(* IEC 61131-3 sources: daoli-st-library/DL_Algo (part 14) *)

(* ---- FB_DL_GainSchedPid.st ---- *)
(*
  组件名 Component   : FB_DL_GainSchedPid
  子库 Sublibrary    : DL_Algo
  版本 Version       : 1.0.0
  兼容性 Platform    : CODESYS 3.5 / TwinCAT 3 / 汇川 InoProShop / Machine Expert（仅 Standard.library）
  功能 Function      : 增益调度 PID（T0 标准语义件）：
                       1) 按调度变量 fSchedX 在断点表 afSchedX 上分区线性插值 Kc/Ti/Td 参数集；
                       2) 区间过渡加权平滑：插值参数经一阶惯性（tGainSmooth）再入 PID 核，
                          防分区切换瞬间增益阶跃引起执行器冲击；
                       3) 内嵌并行式 PID 核（P + I + D），积分钳位抗饱和，输出限幅；
                       4) 组态闸：断点数域 [2, 8]、断点严格递增、Ti > 0、增益非有限 → 故障锁存。
  边界 Boundary      : ① 本件只出控制量 fCtrlOut，不写物理 IO（由上层适配层承载）；
                       ② 除法防护：Ti 下限 1.0E-6 s、调度跨度判零、tCycle 域闸后再进算式；
                       ③ 非有限值（NaN 自反 + 无穷差值自减）判组态/输入非法，锁存安全侧；
                       ④ 调度变量越断点表两端时取端点参数（钳位外推禁止）；
                       ⑤ 故障锁存解除唯一路径 = bReset 上升沿（输入引脚，恒可达）；
                       ⑥ 无全局变量引用、无外部变量声明、无物理地址寻址。
  依赖 Depends       : Standard.library（R_TRIG）
  溯源 Origin        : IEC 61131-3 标准语义的道莅防御性实现（增益调度 + 并行 PID 均为
                       公开标准控制语义，T0 口径；参考 t2-5-modpid 参数域划分，零代码行复制）
  码位 Code          : 16#02_3_8C
  码表 Error codes（Algo 格 02_3_8C，单轨：故障 0x038C / 信息 0x028C）:
    16#0002_038C 故障级：组态非法（断点数越 [2,8] / 断点非严格递增 / Ti <= 0 /
                 参数非有限 / tCycle <= T#0S），锁存至 bReset 上升沿
    16#0002_028C 信息级：调度变量越端点已钳位（不置 bError，每拍瞬时口径）
  修订历史 Revision  :
    2026-11-19  v1.0.0  R44 首版（批次 1 · 序号 2）
*)

TYPE E_DL_GspState :
(
    eIdle  := 0,    // 空闲：未使能，出口冻结 / Idle, outputs frozen
    eRun   := 10,   // 运行：调度插值 + PID 闭环 / Running, scheduling plus PID loop
    eFault := 90    // 故障：组态非法锁存 / Fault, configuration latched
);
END_TYPE

FUNCTION_BLOCK FB_DL_GainSchedPid
VAR_INPUT
    bEnable    : BOOL;                        // 使能，FALSE 时出口冻结 [-] / Enable
    bReset     : BOOL;                        // 上升沿清故障锁存 [-] / Reset edge
    fSetpoint  : REAL;                        // 设定值 [工程单位] / Setpoint
    fFeedback  : REAL;                        // 反馈值 [工程单位] / Feedback
    fSchedX    : REAL;                        // 调度变量（工况量）[工程单位] / Scheduling variable
    afSchedX   : ARRAY[1..8] OF REAL;         // 断点表（须严格递增）[工程单位] / Scheduling breakpoints
    afKc       : ARRAY[1..8] OF REAL;         // 各断点比例增益 [无量纲] / Kc per breakpoint
    afTi       : ARRAY[1..8] OF REAL;         // 各断点积分时间 [秒] / Ti per breakpoint
    afTd       : ARRAY[1..8] OF REAL;         // 各断点微分时间 [秒] / Td per breakpoint
    nPtCount   : INT := 2;                    // 断点数 [个]，域 2..8 / Breakpoint count
    tGainSmooth: TIME := T#1S;                // 增益平滑惯性时间 [毫秒] / Gain smoothing lag
    fOutMin    : REAL := 0.0;                 // 输出下限 [%] / Output floor
    fOutMax    : REAL := 100.0;               // 输出上限 [%] / Output ceiling
    tCycle     : TIME := T#10MS;              // 扫描周期 [毫秒]，须与实际一致 / Scan cycle time
    bResetInt  : BOOL := TRUE;                // 使能下降沿后积分复归 [-] / Reset integral on disable
END_VAR
VAR_OUTPUT
    fCtrlOut   : REAL;                        // 控制量输出 [%] / Control output
    fKcUse     : REAL;                        // 平滑后生效比例增益 [无量纲] / Effective Kc
    fTiUse     : REAL;                        // 平滑后生效积分时间 [秒] / Effective Ti
    fTdUse     : REAL;                        // 平滑后生效微分时间 [秒] / Effective Td
    bError     : BOOL;                        // 故障锁存标志 [-] / Fault latch flag
    uErrId     : UDINT;                       // 事件码，0 = 无事件 / Event code
    eState     : E_DL_GspState;               // 状态出口，段尾单点映射 / State outlet
END_VAR
VAR
    rtReset    : R_TRIG;                      // 复位沿实例，段 0 每拍无条件刷新 / Reset edge
    _eState    : E_DL_GspState := E_DL_GspState.eIdle;  // 内部相位（CASE 唯一写入目标） / Internal phase
    _fErr      : REAL;                        // 偏差 [工程单位] / Error
    _fP        : REAL;                        // 比例项 [%] / Proportional term
    _fI        : REAL;                        // 积分项 [%] / Integral term
    _fD        : REAL;                        // 微分项 [%] / Derivative term
    _fErrPrev  : REAL;                        // 上拍偏差快照 [工程单位] / Previous error
    _fKcRaw    : REAL;                        // 插值比例增益 [无量纲] / Interpolated Kc
    _fTiRaw    : REAL;                        // 插值积分时间 [秒] / Interpolated Ti
    _fTdRaw    : REAL;                        // 插值微分时间 [秒] / Interpolated Td
    _fSeg      : REAL;                        // 插值段权重 [无量纲] / Interpolation weight
    _fCyS      : REAL;                        // 扫描周期秒值 [秒] / Cycle time in seconds
    _fSmK      : REAL;                        // 平滑系数 [无量纲] / Smoothing coefficient
    _nIdx      : INT;                         // 断点搜索索引 [-] / Breakpoint search index
    _bCfgBad   : BOOL;                        // 组态非法当拍量 [-] / Config illegal flag
    _bSchedClp : BOOL;                        // 调度钳位当拍量 [-] / Schedule clamped flag
    _fTiSafe   : REAL;                        // 积分时间安全值 [秒] / Ti safety value
END_VAR
VAR CONSTANT
    DL_PT_MAX  : INT   := 8;                  // 断点数上限，与数组维度一致 [个] / Breakpoint ceiling
    DL_PT_MIN  : INT   := 2;                  // 断点数下限 [个] / Breakpoint floor
    DL_MS_PER_S: REAL  := 1000.0;             // 毫秒 → 秒换算系数 [毫秒/秒] / Milliseconds per second
    DL_TI_MIN  : REAL  := 1.0E-6;             // 积分时间下限 [秒] / Ti floor
    DL_ABS_MAX : REAL  := 1.0E30;             // 有限值判定上界 [工程单位] / Finite value bound
    DL_EPS     : REAL  := 1.0E-9;             // 跨度判零容差 [工程单位] / Zero span tolerance
    DL_ZERO    : REAL  := 0.0;                // 零常量 [工程单位] / Zero constant
    DL_ONE     : REAL  := 1.0;                // 单位常量 [无量纲] / Unity constant
    DL_NO_TIME : TIME  := T#0S;               // 零时长哨兵 [毫秒] / Zero time sentinel
END_VAR

(* —— 段 0｜沿实例每拍无条件刷新（禁置于 IF/CASE 内） —— *)
rtReset(CLK := bReset);

(* —— 段 1｜瞬时量预清零（锁存量 _eState/积分项不入清单，禁同拍抹除） —— *)
_bCfgBad   := FALSE;
_bSchedClp := FALSE;
uErrId     := 16#0000_0000;

(* —— 段 2｜复位沿：故障一次性清干净，相位回空闲 —— *)
IF rtReset.Q THEN
    _eState  := E_DL_GspState.eIdle;
    _fI      := DL_ZERO;
    _fErrPrev:= DL_ZERO;
END_IF

(* —— 段 3｜周期换算与组态闸（覆盖全部参与换算引脚） —— *)
_fCyS := TIME_TO_REAL(tCycle) / DL_MS_PER_S;    // 毫秒 → 秒（TIME_TO_REAL 标准转换）
IF (tCycle = DL_NO_TIME) OR (nPtCount < DL_PT_MIN) OR (nPtCount > DL_PT_MAX) THEN
    _bCfgBad := TRUE;
END_IF
IF NOT _bCfgBad THEN
    _nIdx := 1;
    WHILE (_nIdx < nPtCount) AND (NOT _bCfgBad) DO
        IF (afSchedX[_nIdx] <> afSchedX[_nIdx]) OR (afKc[_nIdx] <> afKc[_nIdx])
           OR (afTi[_nIdx] <> afTi[_nIdx]) OR (afTd[_nIdx] <> afTd[_nIdx])
           OR (afSchedX[_nIdx + 1] <= afSchedX[_nIdx]) OR (afTi[_nIdx] <= DL_EPS)
           OR (afTi[_nIdx] > DL_ABS_MAX) THEN
            _bCfgBad := TRUE;               // 断点非递增 / 参数非有限 / Ti 无效
        END_IF
        _nIdx := _nIdx + 1;
    END_WHILE;
END_IF

(* —— 段 4｜主状态机：三态全覆盖 + ELSE 兜底 —— *)
CASE _eState OF

E_DL_GspState.eIdle:
    IF bEnable AND (NOT _bCfgBad) THEN
        _fI       := DL_ZERO;               // 入运行相前积分清零
        _fErrPrev := DL_ZERO;
        _eState   := E_DL_GspState.eRun;
    ELSIF bEnable AND _bCfgBad THEN
        bError    := TRUE;                  // 故障级配对置位（R45）
        uErrId    := 16#0002_038C;          // 组态非法锁存
        _eState   := E_DL_GspState.eFault;
    END_IF

E_DL_GspState.eRun:
    IF NOT bEnable THEN
        IF bResetInt THEN
            _fI := DL_ZERO;                 // 使能撤销按组态复归积分
        END_IF
        _eState := E_DL_GspState.eIdle;
    ELSE
        (* 调度插值：越端点钳位取端点参数并留信息码 *)
        IF fSchedX <= afSchedX[1] THEN
            _nIdx      := 1;
            _fSeg      := DL_ZERO;
            _bSchedClp := TRUE;
        ELSIF fSchedX >= afSchedX[nPtCount] THEN
            _nIdx      := nPtCount - 1;
            _fSeg      := DL_ONE;
            _bSchedClp := TRUE;
        ELSE
            _nIdx := 1;
            WHILE (_nIdx < nPtCount) AND (fSchedX >= afSchedX[_nIdx + 1]) DO
                _nIdx := _nIdx + 1;         // 断点严格递增已由组态闸保证
            END_WHILE;
            _fSeg := (fSchedX - afSchedX[_nIdx]) / (afSchedX[_nIdx + 1] - afSchedX[_nIdx]);
        END_IF
        _fKcRaw := afKc[_nIdx] + _fSeg * (afKc[_nIdx + 1] - afKc[_nIdx]);
        _fTiRaw := afTi[_nIdx] + _fSeg * (afTi[_nIdx + 1] - afTi[_nIdx]);
        _fTdRaw := afTd[_nIdx] + _fSeg * (afTd[_nIdx + 1] - afTd[_nIdx]);

        (* 一阶惯性平滑：系数域闸后加权，tGainSmooth 为零时直通 *)
        IF tGainSmooth <= DL_NO_TIME THEN
            _fSmK := DL_ONE;
        ELSE
            _fSmK := _fCyS / (_fCyS + TIME_TO_REAL(tGainSmooth) / DL_MS_PER_S);
        END_IF
        fKcUse := fKcUse + _fSmK * (_fKcRaw - fKcUse);
        fTiUse := fTiUse + _fSmK * (_fTiRaw - fTiUse);
        fTdUse := fTdUse + _fSmK * (_fTdRaw - fTdUse);
        IF _bSchedClp THEN
            uErrId := 16#0002_028C;         // 信息级：调度钳位（瞬时口径）
        END_IF

        (* PID 核：并行式，积分钳位抗饱和 *)
        _fErr := fSetpoint - fFeedback;
        _fP   := fKcUse * _fErr;
        _fTiSafe := MAX(fTiUse, DL_TI_MIN); // 积分时间下限护栏（除零前置）
        _fI := _fI + (fKcUse / _fTiSafe) * _fErr * _fCyS;
        _fD := (fKcUse * fTdUse / _fCyS) * (_fErr - _fErrPrev);
        fCtrlOut := _fP + _fI + _fD;
        IF fCtrlOut > fOutMax THEN
            fCtrlOut := fOutMax;
            _fI := _fI - (fKcUse / _fTiSafe) * _fErr * _fCyS;   // 上饱和积分回退
        ELSIF fCtrlOut < fOutMin THEN
            fCtrlOut := fOutMin;
            _fI := _fI - (fKcUse / _fTiSafe) * _fErr * _fCyS;   // 下饱和积分回退
        END_IF
        _fErrPrev := _fErr;
    END_IF

E_DL_GspState.eFault:
    ;                                   // 故障相驻留：出口冻结，只认复位沿（段 2 承载迁出）

ELSE
    bError := TRUE;                     // 兜底：非法相位锁存
    uErrId := 16#0002_038C;
    _eState := E_DL_GspState.eFault;
END_CASE

(* —— 段 5｜状态出口单点映射 —— *)
eState := _eState;
END_FUNCTION_BLOCK

(* ---- FB_DL_GainScheduler.st ---- *)
(*
    FB_DL_GainScheduler —— 分段增益调度
    ------------------------------------------------------------------
    分类      : DL_Algo / Control
    前缀      : FB_DL_
    版本      : 1.0.0
    溯源      : T2-5 Mod_PID（只借「参数域约束」的组织方式；源矩阵判定其参数域已取尽，
                仅剩「分段 / 手自动」这类手册细节，本件即分段这一侧的收口件）；
                迟滞判据、状态化输出、码位与分级 100% 自有；
                clean-room 重写，未复制任何闭源厂商源码，参考实现仅限 MIT/Apache 许可
    平台      : 纯 IEC 61131-3，CODESYS V3.5+ / TwinCAT 3 / InoProShop 通用
    作者      : 道莅代码库 · PLC编程专家（R18）
    ------------------------------------------------------------------
    功能说明  : 按调度变量（温度 / 流量 / 负载率）落在哪个断点区间，输出该段的一组
                Kp / Ki / Kd，解决「升温段要大 P、保温段要强 I」的分段整定需求；
                核心防御是边界迟滞：升段要越过「断点 + 迟滞半宽」，降段要跌破
                「断点 - 迟滞半宽」，杜绝边界抖动导致增益每拍来回跳；
                复位沿优先于定位，断点表严格递增在校验层一次性拦截；
                职责边界：本件只输出增益，不实现积分，也不做无扰切换——无扰由
                FB_DL_BumplessTransfer 与 PID 侧承担，避免与级联 PID 抢职责。
    错误码    : 16#0002_2301 调度变量非有限或变化被迟滞带抑制（保持当前段）——信息级，不置故障
                16#0002_2302 预留禁用（信息级，不得挪用）
                16#0002_2310 断点表非严格递增（非法组态）——故障级，输出保持末次并置故障
                16#0002_2311 段数越界（不在 2~4）——故障级，输出全 0 且不索引数组
                16#0002_2312 预留禁用（故障级，不得挪用）
    码位总账  : 16#0002_2301 用 / 16#0002_2302 预留 ｜ 16#0002_2310 用 / 16#0002_2311 用 / 16#0002_2312 预留
    状态机    : 无 CASE，段号由 uSeg 一个整数承载，非法状态由段数闸拦截，不可能出现
    采样约定  : fbTrigReset 在本体首部无条件刷新；本件无时间量，切换判定与任务周期无关，
                bSwitched 为单周期脉冲（每拍先清后置）。
    修订记录  : 2026-11-16 v1.0.0 首次入库（R18）
*)
FUNCTION_BLOCK FB_DL_GainScheduler
VAR_INPUT
    bEnable       : BOOL;                      // 使能，FALSE 输出保持末次并冻结段号 / enable, FALSE holds the last gains and freezes the segment
    bReset        : BOOL;                      // 复位，上升沿强制回到段 0 并清切换沿 / reset, rising edge forces segment zero and clears the switch pulse
    fScheduleVar  : REAL := 0.0;               // 调度变量（如温度）[用户单位] / scheduling variable such as temperature [user unit]
    afBreakpoint  : ARRAY[0..3] OF REAL;       // 分段上界断点，有效项 0~uSegCount-2，必须严格递增 [用户单位] / segment upper breakpoints, valid items 0~uSegCount-2, strictly increasing [user unit]
    afKp          : ARRAY[0..3] OF REAL;       // 各段比例增益 [无量纲] / proportional gain per segment [dimensionless]
    afKi          : ARRAY[0..3] OF REAL;       // 各段积分增益 [1/s] / integral gain per segment [1/s]
    afKd          : ARRAY[0..3] OF REAL;       // 各段微分增益 [s] / derivative gain per segment [s]
    uSegCount     : UINT := 2;                 // 段数 [段]，范围 2~4 / segment count [seg], range 2~4
    fHysteresis   : REAL := 0.5;               // 段边界迟滞带半宽 [用户单位]，范围 0.0~100.0，0 = 无迟滞 / half width of the boundary hysteresis band [user unit], range 0.0~100.0, 0 = none
END_VAR
VAR_OUTPUT
    fKp         : REAL;                        // 当前段比例增益 [无量纲] / proportional gain of the active segment [dimensionless]
    fKi         : REAL;                        // 当前段积分增益 [1/s] / integral gain of the active segment [1/s]
    fKd         : REAL;                        // 当前段微分增益 [s] / derivative gain of the active segment [s]
    uActiveSeg  : UINT;                        // 当前段号 0~3 [段] / active segment index 0~3 [seg]
    bSwitched   : BOOL;                        // 段切换单周期脉冲 / single-cycle segment switch pulse
    uSwitchCnt  : UDINT;                       // 累计切换次数，抖动监视用，饱和计数 [次] / accumulated switch count for chatter monitoring, saturating [times]
    eErr        : UDINT;                       // 错误码，0=正常 / error id, 0=ok
    bError      : BOOL;                        // 故障标志，eErr 为故障级时 TRUE / error flag, TRUE on fault-level eErr
END_VAR
VAR
    fbTrigReset : R_TRIG;                      // 复位沿检测实例，本体首部无条件刷新 / reset edge instance, refreshed unconditionally
    bInit       : BOOL := FALSE;               // 首扫标志，初值 FALSE，判据 NOT bInit / first-scan flag, initial FALSE, tested with NOT
    uSeg        : UINT;                        // 内部当前段号 [段] / internal active segment index [seg]
    uIdx        : UINT;                        // 断点遍历游标 [段] / breakpoint traversal cursor [seg]
    fHystEff    : REAL;                        // 生效迟滞半宽，钳位后使用 [用户单位] / effective hysteresis half width after clamping [user unit]
    bNonFin     : BOOL;                        // 调度变量非有限判定标志 / scheduling variable non-finite flag
    uSegLast    : UINT;                        // 上一拍段号，用于切换沿判定 [段] / previous cycle segment index for the switch edge [seg]
END_VAR
VAR CONSTANT
    DL_GS_SEG_MAX     : UINT := 4;             // 段数上限 [段] / segment count upper bound [seg]
    DL_GS_SEG_MIN     : UINT := 2;             // 段数下限 [段] / segment count lower bound [seg]
    DL_GS_LAST_IDX    : UINT := 3;             // 增益数组末索引 [段] / last gain array index [seg]
    DL_GS_HYST_MAX    : REAL := 100.0;         // 迟滞半宽上限 [用户单位] / hysteresis half width upper bound [user unit]
    DL_FLOAT_EPS      : REAL := 1.0E-6;        // 浮点判等容差 [用户单位] / float equality tolerance [user unit]
    DL_GS_INF_GUARD   : REAL := 4.0E38;        // 非有限幅值判定阈值 [用户单位] / non-finite magnitude guard [user unit]
    DL_GS_CNT_MAX     : UDINT := 16#FFFF_FFFE; // 切换计数饱和值 [次] / switch counter saturation value [times]
    DL_GS_ZERO        : REAL := 0.0;           // 零值常量，避免裸字面量 [无量纲] / zero constant, avoids a bare literal [dimensionless]
END_VAR

// 段 1｜边沿实例无条件周期刷新（红线：严禁放入条件分支）/ segment 1, unconditional edge refresh
fbTrigReset(CLK := bReset);

// 段 2｜输出与错误状态预置：bSwitched 每拍先清后置 / segment 2, preset outputs and error status
bSwitched := FALSE;                            // 单拍脉冲先清 / clear the single-cycle pulse first
eErr := 0;                                     // 预置无错误 / preset no error
bError := FALSE;                               // 预置无故障 / preset no fault

// 段 3｜首扫初始化（初值 FALSE，判据 NOT bInit）/ segment 3, first-scan initialisation
IF NOT bInit THEN
    uSeg := 0;                                 // 首扫落段 0 / start in segment zero
    uSegLast := 0;                             // 切换沿比较基准清零 / clear the switch edge reference
    uSwitchCnt := 0;                           // 切换计数清零 / clear the switch counter
    bInit := TRUE;                             // 首扫只做一次 / first scan runs once only
END_IF

// 段 4｜使能闸：失能保持末次增益并冻结段号 / segment 4, enable gate holds the last gains
IF NOT bEnable THEN
    uActiveSeg := uSeg;                        // 段号镜像保持 / keep the mirrored segment index
    RETURN;                                    // 失能即出口 / disabled is the exit
END_IF

// 段 5｜段数闸：越界即输出全 0 且不索引数组 / segment 5, segment count gate
IF (uSegCount < DL_GS_SEG_MIN) OR (uSegCount > DL_GS_SEG_MAX) THEN
    eErr := 16#0002_2311;                      // 段数越界故障码 / segment count out of range fault id
    bError := TRUE;                            // 置故障标志 / raise the error flag
    fKp := DL_GS_ZERO;                         // 输出全 0 / zero all gains
    fKi := DL_GS_ZERO;                         // 输出全 0 / zero the integral gain
    fKd := DL_GS_ZERO;                         // 输出全 0 / zero the derivative gain
    uActiveSeg := 0;                           // 段号回 0 / segment index back to zero
    RETURN;                                    // 故障级提前返回 / early return on fault
END_IF

// 段 6｜断点严格递增校验（浮点用大于号，禁用判等）/ segment 6, strict monotonic breakpoint check
FOR uIdx := 1 TO uSegCount - 2 DO
    IF NOT (afBreakpoint[uIdx] > afBreakpoint[uIdx - 1]) THEN
        eErr := 16#0002_2310;                  // 断点非法故障码 / illegal breakpoint fault id
        bError := TRUE;                        // 置故障标志 / raise the error flag
        uActiveSeg := uSeg;                    // 段号保持，输出保持末次 / keep the segment and the last gains
        RETURN;                                // 故障级提前返回 / early return on fault
    END_IF
END_FOR

// 段 7｜迟滞半宽双向钳位（负值视为无迟滞，超上限钳位）/ segment 7, hysteresis half width clamp
fHystEff := MIN(MAX(fHysteresis, DL_GS_ZERO), DL_GS_HYST_MAX); // 双侧钳位 / clamp both sides

// 段 8｜段号上界保护：段表缩短后旧段号可能越界 / segment 8, segment index upper bound protection
IF uSeg > (uSegCount - 1) THEN
    uSeg := uSegCount - 1;                     // 钳到最高段 / clamp to the highest segment
END_IF

// 段 9｜复位沿优先于定位 / segment 9, reset edge has priority over locating
IF fbTrigReset.Q THEN
    uSeg := 0;                                 // 强制回段 0 / force back to segment zero
END_IF

// 段 10｜迟滞定位：一次调用最多跨一段，跨多段交给后续拍 / segment 10, hysteresis locating, one step per cycle
bNonFin := (fScheduleVar <> fScheduleVar)
        OR (fScheduleVar > DL_GS_INF_GUARD)
        OR (fScheduleVar < -DL_GS_INF_GUARD);   // 非有限判定 / non-finite check
IF bNonFin THEN
    eErr := 16#0002_2301;                      // 非有限保持当前段（信息级不置故障）/ non-finite keeps the current segment, info level never raises a fault
ELSIF (NOT fbTrigReset.Q) THEN
    IF (uSeg < (uSegCount - 1)) AND (fScheduleVar > (afBreakpoint[uSeg] + fHystEff)) THEN
        uSeg := uSeg + 1;                      // 升段：必须越过断点加迟滞 / step up only beyond the breakpoint plus hysteresis
    ELSIF (uSeg > 0) AND (fScheduleVar < (afBreakpoint[uSeg - 1] - fHystEff)) THEN
        uSeg := uSeg - 1;                      // 降段：必须跌破断点减迟滞 / step down only below the breakpoint minus hysteresis
    END_IF
END_IF

// 段 11｜切换沿与抖动计数：段号变化才产生单拍脉冲 / segment 11, switch edge and chatter counting
IF uSeg <> uSegLast THEN
    bSwitched := TRUE;                         // 段号变化即置单拍脉冲 / raise the single-cycle pulse on any change
    IF uSwitchCnt < DL_GS_CNT_MAX THEN
        uSwitchCnt := uSwitchCnt + 1;          // 饱和加一，绝不回绕 / saturating increment, never wraps
    END_IF
END_IF
uSegLast := uSeg;                              // 记录本拍段号供下一拍比较 / remember this cycle segment for the next comparison

// 段 12｜增益输出：段号已由段 8 与段 5 双重保证在合法区间 / segment 12, publish the gains
fKp := afKp[uSeg];                             // 段号不超过 3，索引安全 / the segment index never exceeds three, indexing is safe
fKi := afKi[uSeg];                             // 积分增益取本段表值 / integral gain from the active segment row
fKd := afKd[uSeg];                             // 微分增益取本段表值 / derivative gain from the active segment row
uActiveSeg := uSeg;                            // 对外镜像段号 / publish the segment index
END_FUNCTION_BLOCK

(* ---- FB_DL_GapForceSwitchover.st ---- *)
(*==============================================================================
 * 组件名称 (Component)  : FB_DL_GapForceSwitchover
 * 所属子库 (Sublibrary) : DL_Algo
 * 当前版本 (Version)    : 1.0.0
 * 兼容性   (Platform)   : CODESYS 3.5+ / TwinCAT 3 / 汇川 InoProShop / 施耐德 Machine Expert
 *                         仅依赖 Standard.library（TON / R_TRIG / ABS / MAX），零厂商私有库
 * 功能描述 (Function)   : 压装/贴合类工步位置/压力双模式无扰切换：
 *                           eApproach 接近段：位置控趋近 fGapTargetMm，fCmdTrim = 间隙误差
 *                             修调（钳 ±fTrimMaxMm）；
 *                           接触判据：fForceN >= fContactN + 迟滞带 → eContact 过渡态，
 *                             冻结当时修调/速度作为衔接保持值（切换点速度不得突跳），
 *                             保持一个 tHoldXf 衔接窗后必迁出（单过渡态禁驻留，R285）；
 *                           eForceCtl 力控段：力偏差 → fForceTrimPct（钳 ±100%），
 *                             fCmdTrim 置 0；
 *                           tContactTmo 内未判接触 → eFault（eCause=eNoContact）；
 *                           力传感器非有限/超量程 → eFault（eCause=eForceBad）。
 * 接口     (Interface)  : 输入 fPosMm/fVelMmS 轴位姿、fForceN 力（N）、fContactN 接触判据
 *                         （N）、fGapTargetMm 目标间隙（mm）、fForceTargetN 力控目标（N）、
 *                         tContactTmo 接触超时、tHoldXf 衔接窗、fHysN 接触迟滞（N）、
 *                         fTrimMaxMm 修调限幅（mm）、fKpAppPct 接近修调增益（1/mm）、
 *                         fKpForcePct 力控增益（%/N）、fForceMaxN 力量程上限（N）、bReset；
 *                         输出 eMode 五态、fCmdTrim 位置环修调、fForceTrimPct 力环输出
 *                         （%）、eCause 成因、bError。
 * 边界     (Boundary)   : ① **属主边界（写死）：本件只出双模式状态与两侧修调量，不注入
 *                         轴指令、不接管压力环 PID**；修调限速可由上层用
 *                         `FB_DL_RateLimiter` 串联（本件不内嵌，规格依赖声明）。
 *                         ② 五态 CASE + ELSE 兜底 eFault（R6）；切换判据浮点容差比较
 *                         （迟滞带显式写出，禁 = 判等）。
 *                         ③ eContact 为单过渡态：tHoldXf 到时必迁 eForceCtl，禁驻留。
 *                         ④ 衔接保持值（_fTrimHold / _fVelHold）显式写出并在复位沿清零
 *                         （R311 预防：复位沿清状态与保持值）。
 *                         ⑤ 力超量程判据 = fForceN > fForceMaxN 或 fForceN < 0 或非有限
 *                         → eFault eForceBad（成因分码，R190 归因唯一）。
 *                         ⑥ 零全局耦合（无 GVL / VAR_EXTERNAL / 物理地址）。
 * 分工声明 (Scope)      : 与 `FB_DL_CoatingGapMeasure`（测量）与 `FB_DL_RollCompressForce-
 *                         Balance`（力平衡趋势）分工：切换闭环（本件）≠ 测量 ≠ 趋势。
 * 来源标签 (Source Tag) : T2-2 ◐（LBP 压机工艺分类只借"位置段/压力段"分类事实，切换器
 *                         实现自研）
 * 码表     (Codes)      : 本件不占用任何全局数字码位。出口为 ENUM 五态 + LREAL 组 +
 *                         ENUM 成因 + BOOL；数字码位待主控收口阶段统一派号。
 * 红线自检 (Redline)    : R1 ✓ 零 GVL/VAR_EXTERNAL ｜ R2 ✓ 零 %I/%Q/%M ｜ R3 ✓ 纯 IEC 61131-3
 *                         R4 ✓ 迟滞容差 + 非有限/超量程闸 + 修调钳位 ｜ R5 ✓ 声明逐行同行双语注释
 *                         R6 ✓ 五态 CASE 含 ELSE ｜ R7 ✓ 两 TON/一 R_TRIG 段 0 无条件刷新
 * 修订历史 (Revision)   : 2026-11-20  v1.0.0  R48 首版（批次 3 · 序号 13）
 *                         验收向量：接近段间隙误差修调；力越迟滞带 → eContact 冻结保持值；
 *                         衔接窗到 → eForceCtl；tContactTmo 无接触 → eFault eNoContact。
 *==============================================================================*)

TYPE E_DL_GfsMode :
(
    eIdle     := 0,    // 待机 / Idle
    eApproach := 10,   // 接近段（位置控）/ Approach phase, position control
    eContact  := 20,   // 接触过渡态（衔接保持，单过渡禁驻留）/ Contact transition, hold window
    eForceCtl := 30,   // 力控段 / Force control phase
    eFault    := 90    // 故障（等复位）/ Fault, awaiting reset
);
END_TYPE

TYPE E_DL_GfsCause :
(
    eNone       := 0,   // 无异常 / No anomaly
    eNoContact  := 1,   // 接近段超时未判接触 / No contact within timeout
    eForceBad   := 2,   // 力传感器非有限/超量程/负值 / Force sensor bad
    eCfgIllegal := 3,   // 组态非法 / Illegal configuration
    eModeBad    := 4    // 非法模式兜底 / Illegal mode fallback
);
END_TYPE

FUNCTION_BLOCK FB_DL_GapForceSwitchover
VAR_INPUT
    fPosMm      : LREAL := 0.0;    // 轴实际位置 [mm] / Axis actual position [mm]
    fVelMmS     : LREAL := 0.0;    // 轴实际速度 [mm/s] / Axis actual velocity [mm/s]
    fForceN     : LREAL := 0.0;    // 力/压力传感器实测 [N] / Force sensor measurement [N]
    fContactN   : LREAL := 5.0;    // 接触判据力，域 > 0 [N] / Contact force threshold [N]
    fGapTargetMm: LREAL := 0.0;    // 接近段目标间隙 [mm] / Approach target gap [mm]
    fForceTargetN: LREAL := 100.0; // 力控段目标力 [N] / Force-control target [N]
    tContactTmo : TIME := T#10S;   // 接近段接触超时，域 > T#0S [ms] / Contact timeout [ms]
    tHoldXf     : TIME := T#200MS; // eContact 衔接保持窗，域 > T#0S [ms] / Transition hold window [ms]
    fHysN       : LREAL := 0.5;    // 接触判据迟滞带，域 >= 0 [N] / Contact hysteresis band [N]
    fTrimMaxMm  : LREAL := 1.0;    // 位置环修调限幅，域 > 0 [mm] / Position trim limit [mm]
    fKpAppPct   : LREAL := 1.0;    // 接近段修调增益（间隙误差→修调） [1/mm] / Approach trim gain [1/mm]
    fKpForcePct : LREAL := 0.5;    // 力控段增益（力偏差→%） [%/N] / Force-control gain [%/N]
    fForceMaxN  : LREAL := 5000.0; // 力传感器量程上限，域 > fContactN [N] / Force range ceiling [N]
    bReset      : BOOL := FALSE;   // 故障复位，上升沿回 eIdle 并清保持值（R311） [-] / Fault reset, rising edge clears state and holds
END_VAR
VAR_OUTPUT
    eMode        : E_DL_GfsMode;   // 双模式状态出口 [-] / Mode state outlet
    fCmdTrim     : LREAL;          // 位置环速度/位置修调输出（力控段恒 0） [mm] / Position-loop trim outlet [mm]
    fForceTrimPct: LREAL;          // 力环修调输出（接近段恒 0） [%] / Force-loop trim outlet [%]
    eCause       : E_DL_GfsCause;  // 成因出口（锁存回放，R189） / Cause outlet, latched
    bError       : BOOL;           // 故障标志 [-] / Error flag
END_VAR
VAR
    _eMode     : E_DL_GfsMode := E_DL_GfsMode.eIdle;   // 内部状态（CASE 唯一写入目标） / Internal mode
    _eCause    : E_DL_GfsCause := E_DL_GfsCause.eNone; // 成因锁存量 / Latched cause
    _bFault    : BOOL;           // 故障锁存位（解除沿 = bReset 上升沿） / Latched fault bit
    _fTrimHold : LREAL := 0.0;   // 衔接保持值：接触瞬间修调 [mm] / Held trim at contact
    _fVelHold  : LREAL := 0.0;   // 衔接保持值：接触瞬间速度 [mm/s] / Held velocity at contact
    _fForceTrim: LREAL := 0.0;   // 力环修调锁存镜像 [%] / Force trim latch mirror
    _fCmdTrim  : LREAL := 0.0;   // 位置修调锁存镜像 [mm] / Position trim latch mirror
    _bErrScan  : BOOL;           // 力信号病当拍量（触发 eFault 用） / Force bad this scan
    _bNonFin   : BOOL;           // 输入非有限当拍量 [-] / Non-finite input this scan
    _bCfgBad   : BOOL;           // 组态非法当拍量 [-] / Illegal configuration this scan
    tonContactTmo: TON;          // 接近段接触超时定时器，段 0 无条件调用 / Contact timeout timer
    tonHoldXf  : TON;            // 衔接保持窗定时器，段 0 无条件调用 / Transition hold timer
    rtReset    : R_TRIG;         // 复位沿实例，段 0 无条件调用 / Reset edge instance
END_VAR
VAR CONSTANT
    DL_GFS_EPS   : LREAL := 1.0E-6;  // 浮点判零容差 [无量纲] / Float epsilon
    DL_GFS_ZERO  : LREAL := 0.0;     // 非有限差值判零基准 [-] / Non-finite difference zero base
    DL_GFS_PCTMAX: LREAL := 100.0;   // 力环修调行程上限 [%] / Force trim travel ceiling [%]
END_VAR

(* —— 段 0：非有限判 + 组态闸 + 两 TON 一沿无条件周期刷新 —— *)
_bNonFin := (fForceN <> fForceN) OR ((fForceN - fForceN) <> DL_GFS_ZERO)
         OR (fPosMm <> fPosMm) OR (fVelMmS <> fVelMmS);   // 力/位置/速度非有限（R245） / Non-finite force, position, velocity
_bCfgBad := (fContactN <= DL_GFS_ZERO) OR (fForceMaxN <= fContactN)
         OR (tContactTmo <= T#0S) OR (tHoldXf <= T#0S)
         OR (fTrimMaxMm <= DL_GFS_ZERO) OR (fHysN < DL_GFS_ZERO);   // 组态域闸 / Configuration gate
_bErrScan := _bNonFin OR (fForceN > fForceMaxN) OR (fForceN < DL_GFS_ZERO);   // 力信号病（超量程/负值/非有限） / Force signal bad
tonContactTmo(IN := (_eMode = E_DL_GfsMode.eApproach), PT := tContactTmo);   // 接触超时（进接近段计时，出段自复位） / Contact timeout
tonHoldXf(IN := (_eMode = E_DL_GfsMode.eContact), PT := tHoldXf);   // 衔接保持窗（进过渡态计时） / Transition hold window
rtReset(CLK := bReset);                                     // 复位沿，每拍必调 / Reset edge, every scan

(* —— 段 1：组态闸入故障 —— *)
IF _bCfgBad AND (NOT _bFault) THEN
    _bFault := TRUE;                                        // 组态非法锁存 / Latch config fault
    _eCause := E_DL_GfsCause.eCfgIllegal;                   // 归因：组态非法 / Cause: illegal config
    _eMode := E_DL_GfsMode.eFault;                          // 入故障态 / Enter fault
END_IF

(* —— 段 2：迁出链（复位沿：清状态与保持值，R311 预防） —— *)
IF rtReset.Q THEN
    _bFault := FALSE;                                       // 清故障锁存 / Clear fault latch
    _eCause := E_DL_GfsCause.eNone;                         // 清成因 / Clear cause
    _fTrimHold := 0.0;                                      // 清衔接保持修调 / Clear held trim
    _fVelHold := 0.0;                                       // 清衔接保持速度 / Clear held velocity
    _fCmdTrim := 0.0;                                       // 清修调镜像 / Clear trim mirror
    _fForceTrim := 0.0;                                     // 清力环镜像 / Clear force mirror
    _eMode := E_DL_GfsMode.eIdle;                           // 回待机 / Back to idle
END_IF

(* —— 段 3：力信号病 → 故障（成因分码 eForceBad，优先于时序） —— *)
IF _bErrScan AND (NOT _bFault) THEN
    _bFault := TRUE;                                        // 力信号病锁存 / Latch force fault
    _eCause := E_DL_GfsCause.eForceBad;                     // 归因：力传感器病 / Cause: force bad
    _eMode := E_DL_GfsMode.eFault;                          // 入故障态 / Enter fault
END_IF

(* —— 段 4：五态状态机（故障态由迁出链处理） —— *)
IF NOT _bFault THEN
    CASE _eMode OF

    E_DL_GfsMode.eIdle:
        _eMode := E_DL_GfsMode.eApproach;                   // 待机下一拍即入接近段（启动权交上层使能本件调用） / Idle proceeds to approach
        _fCmdTrim := 0.0;                                   // 修调清零起步 / Trim starts at zero

    E_DL_GfsMode.eApproach:
        _fCmdTrim := (fGapTargetMm - fPosMm) * fKpAppPct;   // 接近段修调 = 间隙误差×增益 / Approach trim from gap error
        IF _fCmdTrim > fTrimMaxMm THEN
            _fCmdTrim := fTrimMaxMm;                        // 修调上钳 / Clamp trim high
        ELSIF _fCmdTrim < -fTrimMaxMm THEN
            _fCmdTrim := -fTrimMaxMm;                       // 修调下钳 / Clamp trim low
        END_IF
        IF fForceN >= (fContactN + fHysN) THEN
            _fTrimHold := _fCmdTrim;                        // 接触瞬间冻结修调保持值（无扰衔接，头注释③） / Freeze trim at contact
            _fVelHold := fVelMmS;                           // 冻结接触瞬间速度（防切换突跳） / Freeze velocity at contact
            _fForceTrim := 0.0;                             // 力环修调起步零 / Force trim starts zero
            _eMode := E_DL_GfsMode.eContact;                // 越迟滞带上界：入接触过渡态 / Contact: enter transition
        ELSIF tonContactTmo.Q THEN
            _bFault := TRUE;                                // 超时未接触：故障锁存 / Timeout: latch fault
            _eCause := E_DL_GfsCause.eNoContact;            // 归因：未接触 / Cause: no contact
            _eMode := E_DL_GfsMode.eFault;                  // 入故障态 / Enter fault
        END_IF

    E_DL_GfsMode.eContact:
        _fCmdTrim := _fTrimHold;                            // 衔接窗内保持冻结修调（输出不突跳） / Hold frozen trim in window
        IF tonHoldXf.Q THEN
            _eMode := E_DL_GfsMode.eForceCtl;               // 衔接窗到必迁力控段（单过渡态禁驻留，R285） / Window done forces force phase
        END_IF

    E_DL_GfsMode.eForceCtl:
        _fCmdTrim := 0.0;                                   // 力控段位置修调归零 / Position trim zero in force phase
        _fForceTrim := (fForceTargetN - fForceN) * fKpForcePct;   // 力偏差 → 力环修调 / Force error to trim
        IF _fForceTrim > DL_GFS_PCTMAX THEN
            _fForceTrim := DL_GFS_PCTMAX;                   // 力环上钳 100% / Clamp force trim high
        ELSIF _fForceTrim < -DL_GFS_PCTMAX THEN
            _fForceTrim := -DL_GFS_PCTMAX;                  // 力环下钳 -100% / Clamp force trim low
        END_IF

    E_DL_GfsMode.eFault:
        ;                                                   // 故障态驻留：由段 2 迁出链复位处理 / Held by exit chain in stage 2

    ELSE
        _bFault := TRUE;                                    // 非法模式兜底（R6） / Illegal mode fallback
        _eCause := E_DL_GfsCause.eModeBad;                  // 归因：非法模式 / Cause: illegal mode
        _eMode := E_DL_GfsMode.eFault;                      // 强拉故障态 / Force fault

    END_CASE
END_IF

(* —— 段 5：出口单点映射（名实双出口同源，R191） —— *)
eMode := _eMode;                                            // 模式出口 / Mode outlet
fCmdTrim := _fCmdTrim;                                      // 位置修调出口（故障/待机零） / Position trim outlet
fForceTrimPct := _fForceTrim;                               // 力环修调出口 / Force trim outlet
eCause := _eCause;                                          // 成因出口 / Cause outlet
bError := _bFault OR _bCfgBad OR _bErrScan;                 // 故障标志三源合一 / Error flag
IF bError AND (NOT _bFault) THEN
    _bFault := TRUE;                                        // 当拍病亦锁存（防抖动复归） / Latch scan faults too
END_IF

END_FUNCTION_BLOCK

(* ---- FB_DL_GasDensityComp.st ---- *)
//==============================================================================
// 功能块：FB_DL_GasDensityComp ｜ 中文名称：反应釜气体密度温压补偿
// 所属子库：DL_Algo ｜ 版本：v1.0.0 ｜ 兼容：CODESYS V3.5+ / TwinCAT 3 / 汇川 InoProShop
// 功能描述：理想气体定律温压补偿——由工作温度与绝对压力换算气体密度：
//           rho = p·M / (R·T_K)，M 为介质摩尔质量 [g/mol]，R = 8.314462618
//           [J/(mol·K)]，T_K = T + 273.15。参考态密度 rho_ref 用参考温压
//           同式预计算（诊断出口）。骨架复用 FC_DL_AirDensity 的「域校验
//           + 钳位照算 + 非有限兜底」结构（该件介质常量固定为干空气/
//           水蒸气，反应釜介质摩尔质量可变，故本件以 M 引脚自持实现，
//           不调用该件——Algo 泳道内同口径双实现按 FC_DL_AirDensity 头
//           注释的零依赖纪律执行）。适用域：理想气体偏差可容忍的低压
//           工艺气（N2/Ar/H2/合成气等），近冷凝域给信息级外推提示。
// 开源溯源 (Origin)：道莅原创实现（参考理想气体状态方程与 FC_DL_AirDensity 域校验骨架 分类与参数域）
// 单位表：压力[千帕]（绝对）/ 温度[摄氏度] / 摩尔质量[克每摩尔] /
//         密度[千克每立方米] / 气体常数[J每摩尔开]
// 错误码表：16#0002_3201 信息级（温度/压力域外已钳位照算：温度域
//           [-40, 200] 摄氏度、压力域 [10, 2000] 千帕，不置 bError）/
//           16#0002_3202 信息级（理想气体外推提示：工作点温压比超出
//           参考态 0.5~2 倍温比或 10 倍压比工程带，按理想气体照算，
//           不置 bError）/ 16#0002_3205 预留禁用（不得挪用）/
//           16#0002_3210 故障级（摩尔质量 <= 0 或 > 200，或任一输入
//           非有限，组态非法，置 bError）/ 16#0002_3211 故障级（结果
//           非有限溢出，置 bError——该场景不可由 3210 的组态类判据
//           观测，属数值输出独立域）
// 状态机：E_DL_GasCompState（三态：eIdle=0 / eRun=10 / eFault=99），
//           CASE 含 ELSE 兜底，ELSE 置 3211 并冻结输出零
// 边界行为：① 摩尔质量域外或非有限 → 故障 3210 锁存，bReset 复位；
//           ② 温压域外 → 双侧钳位照算 + 信息 3201（现场宁要标注近似
//           的密度值，不因传感器越量程断链，与骨架件同策略）；
//           ③ 外推带 → 信息 3202 照算；④ 绝对温度下限 233.15 开由温度
//           下限保证，无除零面（T_K 恒正，R 为常量非零）；⑤ 未使能
//           输出冻结为零并 bValid := FALSE；⑥ 安全侧 = 故障/未使能路径
//           输出零密度，禁止残密度进入流量换算下游。
// 修订历史：v1.0.0 2026-11-17 首版（R24 派单 · ROADMAP P2 §670）
//==============================================================================

(*------------------------------------------------------------------------------
 * 枚举: E_DL_GasCompState（归属本功能块，同文件发布，全库唯一定义）
 * 含义: 补偿使能相位，每个成员在 CASE 中有且仅有一个标签。
 *-----------------------------------------------------------------------------*)
TYPE E_DL_GasCompState :
(
    eIdle  := 0,   // 空闲：未使能，输出冻结零 / Idle, not enabled, outputs frozen at zero
    eRun   := 10,  // 运行：使能且组态合法，每拍补偿 / Run, enabled with legal config, compensating per scan
    eFault := 99   // 故障：组态非法/非法状态 / Fault, illegal config or illegal state
);
END_TYPE

FUNCTION_BLOCK FB_DL_GasDensityComp
VAR_INPUT
    fPressKpa    : LREAL := 101.325;        // 工作绝对压力 [千帕]，域 10..2000，域外钳位照算 / Working absolute pressure [kPa], domain 10..2000
    fTempC       : LREAL := 20.0;           // 工作温度 [摄氏度]，域 -40..200，域外钳位照算 / Working temperature [degC], domain -40..200
    fMolarMassG  : LREAL := 28.96;          // 介质摩尔质量 [克每摩尔]，有效域 (0, 200]，空气 28.96 / Medium molar mass [g/mol], valid range (0, 200]
    fPressRefKpa : LREAL := 101.325;        // 参考态绝对压力 [千帕]，须 > 0 / Reference absolute pressure [kPa], must be > 0
    fTempRefC    : LREAL := 20.0;           // 参考态温度 [摄氏度]，须 > -273.15 / Reference temperature [degC], must be above absolute zero
    bEnable      : BOOL;                    // 补偿使能 [—] / Compensation enable
    bReset       : BOOL;                    // 故障复位 [—]，上升沿清组态锁存 / Fault reset, rising edge clears the config latch
END_VAR
VAR_OUTPUT
    fRhoKgM3     : LREAL;                   // 补偿密度 [千克每立方米] / Compensated density [kg/m3]
    fRhoRefKgM3  : LREAL;                   // 参考态密度（诊断出口）[千克每立方米] / Reference density, diagnostics outlet [kg/m3]
    eState       : E_DL_GasCompState;       // 补偿相位 [—] / Compensation phase
    eErr         : UDINT;                   // 错误码，0 = 无错，码位 16#0002_3201 起信息级、16#0002_3210 起故障级（分带见错误码表） / Error code, 0 = no error, band info/fault per the code table
    bError       : BOOL;                    // 故障级标志，仅故障级错误置位 / Fault-class flag, set only on fault-level codes
    bValid       : BOOL;                    // 输出可用标志 / Outputs usable flag
END_VAR
VAR
    _eState      : E_DL_GasCompState := E_DL_GasCompState.eIdle; // 当前相位 / Current phase
    _bParamBad   : BOOL;                    // 摩尔质量/参考态组态非法锁存 / Illegal molar mass or reference config latch
    _bInfoClamp  : BOOL;                    // 温压钳位信息当拍标志 / Temperature or pressure clamp info flag of this scan
    _bInfoExtrap : BOOL;                    // 外推带信息当拍标志 / Extrapolation-band info flag of this scan
    _fTUse       : LREAL;                   // 生效工作温度（已钳位）[摄氏度] / Effective working temperature, clamped
    _fPUse       : LREAL;                   // 生效工作压力（已钳位）[千帕] / Effective working pressure, clamped
    _fTKelvin    : LREAL;                   // 工作绝对温度 [开] / Working absolute temperature [K]
    _fTRefKelvin : LREAL;                   // 参考绝对温度 [开] / Reference absolute temperature [K]
    _bInit       : BOOL := FALSE;           // 首扫标志，初值 FALSE 取非判定 / First-scan flag, tested negated
    _bIllegal    : BOOL;                    // 非法状态标志 / Illegal state flag
END_VAR
VAR CONSTANT
    DL_GDC_R_UNIV  : LREAL := 8.314462618;  // 通用气体常数 [焦耳每摩尔开] / Universal gas constant [J/(mol K)]
    DL_GDC_KELVIN  : LREAL := 273.15;       // 摄氏转开尔文偏移 [开] / Celsius to Kelvin offset [K]
    DL_GDC_T_MIN   : LREAL := -40.0;        // 工作温度域下限 [摄氏度] / Working temperature domain floor [degC]
    DL_GDC_T_MAX   : LREAL := 200.0;        // 工作温度域上限 [摄氏度] / Working temperature domain ceiling [degC]
    DL_GDC_P_MIN   : LREAL := 10.0;         // 工作压力域下限 [千帕] / Working pressure domain floor [kPa]
    DL_GDC_P_MAX   : LREAL := 2000.0;       // 工作压力域上限 [千帕] / Working pressure domain ceiling [kPa]
    DL_GDC_M_MAX   : LREAL := 200.0;        // 摩尔质量域上限 [克每摩尔] / Molar mass domain ceiling [g/mol]
    DL_GDC_MRATIO  : LREAL := 10.0;         // 外推带压比门限 [倍] / Extrapolation pressure-ratio threshold [ratio]
    DL_GDC_TRATIO  : LREAL := 2.0;          // 外推带温比门限（双侧 0.5~2）[倍] / Extrapolation temperature-ratio threshold [ratio]
    DL_GDC_EPS     : LREAL := 1.0E-6;       // 浮点判零容差 [混合] / Float zero tolerance
    DL_GDC_INF     : LREAL := 1.7976931348623157E308; // LREAL 幅值上限 / LREAL magnitude ceiling
    DL_GDC_ZERO    : LREAL := 0.0;          // 零值常量，避免裸字面量 [混合] / Zero constant, avoids a bare literal
END_VAR

(*------------------------------------------------------------------------------
 * 段 1｜每拍预置：输出安全侧清零，单拍标志预清零
 *      Outputs cleared fail-safe first, one-shot flags pre-cleared
 *-----------------------------------------------------------------------------*)
fRhoKgM3    := DL_GDC_ZERO;              // 补偿密度先清（安全侧） / Compensated density cleared first
fRhoRefKgM3 := DL_GDC_ZERO;              // 参考密度先清 / Reference density cleared first
eErr   := 16#0000_0000;                  // 错误码每拍重算 / Error code recomputed
bError := FALSE;                         // 故障标志每拍重算 / Fault flag recomputed
bValid := FALSE;                         // 可用标志每拍重算 / Usable flag recomputed
_bInfoClamp  := FALSE;                   // 钳位信息预清零 / Clamp info pre-cleared
_bInfoExtrap := FALSE;                   // 外推信息预清零 / Extrapolation info pre-cleared
_bIllegal    := FALSE;                   // 非法状态预清零 / Illegal flag pre-cleared

(*------------------------------------------------------------------------------
 * 段 2｜首扫初始化
 *      First-scan initialisation
 *-----------------------------------------------------------------------------*)
IF NOT _bInit THEN
    _eState    := E_DL_GasCompState.eIdle; // 相位空闲起步 / Phase starts idle
    _bParamBad := FALSE;                   // 组态锁存清零 / Config latch cleared
    _bInit     := TRUE;                    // 首扫只做一次 / The first scan runs once
END_IF

(*------------------------------------------------------------------------------
 * 段 3｜组态防御闸：非有限（R79）+ 摩尔质量/参考态物理域
 *      Configuration defense gates: non-finite plus physical domains
 *-----------------------------------------------------------------------------*)
IF (fPressKpa <> fPressKpa) OR (ABS(fPressKpa) > DL_GDC_INF)
   OR (fTempC <> fTempC) OR (ABS(fTempC) > DL_GDC_INF)
   OR (fMolarMassG <> fMolarMassG) OR (ABS(fMolarMassG) > DL_GDC_INF)
   OR (fPressRefKpa <> fPressRefKpa) OR (ABS(fPressRefKpa) > DL_GDC_INF)
   OR (fTempRefC <> fTempRefC) OR (ABS(fTempRefC) > DL_GDC_INF) THEN
    _bParamBad := TRUE;                    // 非有限归组态非法锁存 / Non-finite folded into the config fault latch
END_IF
IF (NOT _bParamBad)
   AND ((fMolarMassG <= DL_GDC_EPS) OR (fMolarMassG > DL_GDC_M_MAX)
        OR (fPressRefKpa <= DL_GDC_EPS) OR (fTempRefC <= (-DL_GDC_KELVIN + 1.0))) THEN
    _bParamBad := TRUE;                    // 摩尔质量/参考态组态非法锁存 / Molar mass or reference config latched
END_IF
IF bReset THEN
    _bParamBad := FALSE;                   // 复位清组态锁存 / Reset clears the config latch
END_IF

(*------------------------------------------------------------------------------
 * 段 4｜相位机（CASE 含 ELSE 兜底；未使能/异常一律落故障态全零）
 *      Phase machine with ELSE fallback, not-enabled or anomaly to fault
 *-----------------------------------------------------------------------------*)
IF (NOT bEnable) OR _bParamBad THEN
    _eState := E_DL_GasCompState.eFault;   // 未使能或组态非法转故障态（全零） / Not enabled or illegal config, fault with zeros
ELSE
CASE _eState OF

    E_DL_GasCompState.eIdle:               // 空闲：使能即进运行
        IF bEnable THEN
            _eState := E_DL_GasCompState.eRun; // 进运行 / To run
        END_IF

    E_DL_GasCompState.eRun:                // 运行：每拍补偿（段 5 执行）
        IF NOT bEnable THEN
            _eState := E_DL_GasCompState.eFault; // 使能撤销转故障态（全零） / Enable dropped, fault with zeros
        END_IF

    E_DL_GasCompState.eFault:              // 故障：使能且复位沿回运行
        IF bEnable AND (NOT _bParamBad) THEN
            _eState := E_DL_GasCompState.eRun; // 回运行 / Back to run
        END_IF

    ELSE                                   // 非法状态兜底（R21：CASE 必带 ELSE）
        _bIllegal := TRUE;                 // 标记非法状态 / Flag the illegal state
        _eState   := E_DL_GasCompState.eFault; // 回故障态（全零） / Back to fault, zeros
END_CASE
END_IF

(*------------------------------------------------------------------------------
 * 段 5｜补偿计算（仅运行态）：域钳位照算 + 外推带提示 + 理想气体定律
 *      Compensation in the run phase: clamp-and-continue plus ideal-gas law
 *-----------------------------------------------------------------------------*)
IF _eState = E_DL_GasCompState.eRun THEN
    _fTUse := fTempC;                      // 工作温度生效 / Working temperature applied
    IF (_fTUse < DL_GDC_T_MIN) OR (_fTUse > DL_GDC_T_MAX) THEN
        _fTUse := MIN(MAX(_fTUse, DL_GDC_T_MIN), DL_GDC_T_MAX); // 温度双侧钳位 / Two-sided temperature clamp
        _bInfoClamp := TRUE;               // 钳位信息置位 / Clamp info raised
    END_IF
    _fPUse := fPressKpa;                   // 工作压力生效 / Working pressure applied
    IF (_fPUse < DL_GDC_P_MIN) OR (_fPUse > DL_GDC_P_MAX) THEN
        _fPUse := MIN(MAX(_fPUse, DL_GDC_P_MIN), DL_GDC_P_MAX); // 压力双侧钳位 / Two-sided pressure clamp
        _bInfoClamp := TRUE;               // 钳位信息置位 / Clamp info raised
    END_IF
    _fTKelvin    := _fTUse + DL_GDC_KELVIN;     // 工作绝对温度 [开]，下限 233.15 恒正 / Working Kelvin, floor 233.15, always positive
    _fTRefKelvin := fTempRefC + DL_GDC_KELVIN;  // 参考绝对温度 [开] / Reference Kelvin
    fRhoKgM3 := (_fPUse * 1000.0) * (fMolarMassG / 1000.0) / (DL_GDC_R_UNIV * _fTKelvin); // 理想气体密度 [千克每立方米]，分母恒正 / Ideal-gas density, denominator always positive
    fRhoRefKgM3 := (fPressRefKpa * 1000.0) * (fMolarMassG / 1000.0) / (DL_GDC_R_UNIV * _fTRefKelvin); // 参考态密度 [千克每立方米] / Reference density
    IF (_fPUse > DL_GDC_MRATIO * fPressRefKpa)
       OR (_fTKelvin < (0.5 * _fTRefKelvin)) OR (_fTKelvin > (DL_GDC_TRATIO * _fTRefKelvin)) THEN
        _bInfoExtrap := TRUE;              // 理想气体外推带提示（照算） / Extrapolation-band notice, computed as-is
    END_IF
END_IF

(*------------------------------------------------------------------------------
 * 段 6｜码位出口与放行（故障级码 3 行内置 bError，R45/R101 配对）
 *      Code outlet and release, fault codes paired with bError
 *-----------------------------------------------------------------------------*)
IF _bIllegal THEN
    eErr   := 16#0002_3211;                // 故障级：状态机兜底（结果域） / Fault: state machine fallback
    bError := TRUE;                        // 置故障标志 / Raise the fault flag
ELSIF _bParamBad THEN
    eErr   := 16#0002_3210;                // 故障级：组态非法 / Fault: illegal configuration
    bError := TRUE;                        // 置故障标志 / Raise the fault flag
ELSIF _bInfoClamp THEN
    eErr := 16#0002_3201;                  // 信息级：温压域外已钳位照算 / Info: clamped, computed as-is
ELSIF _bInfoExtrap THEN
    eErr := 16#0002_3202;                  // 信息级：理想气体外推带照算 / Info: extrapolation band, computed as-is
END_IF

bValid := (NOT bError) AND (_eState = E_DL_GasCompState.eRun); // 仅运行态放行 / Usable only in the run phase
eState := _eState;                       // 相位出口 / Phase outlet
END_FUNCTION_BLOCK

(* ---- FB_DL_GatedUpdateFilter.st ---- *)
(*==============================================================================
 * 组件名称 (Component)  : FB_DL_GatedUpdateFilter
 * 所属子库 (Sublibrary) : DL_Algo
 * 当前版本 (Version)    : 1.0.0
 * 兼容性   (Platform)   : CODESYS 3.5+ / TwinCAT 3 / 汇川 InoProShop / 施耐德 Machine Expert
 *                         仅依赖 Standard.library（TON），零厂商私有库
 * 功能描述 (Function)   : 门控更新滤波：**仅在允许窗口内采样，窗口外保持上次值**。
 *                         与低通 / 限速不同，本件不做任何数值整形，只决定「这一拍要不要采纳」，
 *                         因此阶跃与斜率在窗口内原样通过（无失真、无滞后）。
 *                         典型用途：剔除运动段/换型段的动态值、只在静止窗口内采重量、
 *                         只在保压阶段记录压力稳态值。
 *                         窗口外持续时长用 TON 累计；超过 tMaxHold 置 bStale=TRUE（信息级），
 *                         提示上游「数据已陈旧」，但**输出仍保持**（保持语义不变）。
 *                         恢复路径：bGate 重新为 TRUE 即回到新鲜；故障态由 bEnable 跌落或 bReset 解除。
 * 接口     (Interface)  : 输入 bEnable 使能、bReset 复位到当前输入、fIn 采样输入 [EU]、
 *                         bGate 窗口使能（TRUE = 本拍采纳）、tMaxHold 允许的最大保持时长 [s]；
 *                         输出 fOut 输出值 [EU]、bStale 数据是否陈旧、tHeldElapsed 已保持时长 [s]、
 *                         bValid 输出有效、bError、uErrorId。
 * 边界     (Boundary)   : ① 属主边界：只做门控与保持，不做平滑、不做离群剔除（另件）。
 *                         ② 非有限输入防御：窗口内（bGate=TRUE）遇非有限值 → 故障态 16#0006_0002，
 *                         输出冻结；窗口外（bGate=FALSE）不读取 fIn，故非有限值不判故障
 *                         （这是本件的语义：窗口外输入无意义）。
 *                         ③ tMaxHold < 0 钳到 T#0S 并置信息码 16#0006_0001；T#0S 表示不判陈旧
 *                         （bStale 恒 FALSE，TON 的 Q 仍按 PT=0 立即为真，故显式屏蔽）。
 *                         ④ **TON 无条件每周期调用**（R7），位于 CASE 之外。
 *                         ⑤ 零全局耦合（无 GVL / VAR_EXTERNAL / 物理地址）。
 * 分工声明 (Scope)      : 与 `FB_DL_HoldLastGoodFilter` 分工：坏值（判据失效）保持归那件、
 *                         时间窗门控归本件；与 `FB_DL_PeakHoldFilter` 分工：峰值保持归那件。
 * 来源标签 (Source Tag) : 原创实现（无外部代码引入）
 * 码表     (Codes)      : 16#0006_0000 无故障 / 16#0006_0001 保持时长非法已钳位（信息级）/
 *                         16#0006_0002 窗口内输入非有限（故障级）/ 16#0006_0005 非法状态（故障级）。
 * 红线自检 (Redline)    : R1 ✓ 零 GVL/VAR_EXTERNAL ｜ R2 ✓ 零 %I/%Q/%M ｜ R3 ✓ 纯 IEC 61131-3
 *                         R4 ✓ 非有限拒绝（仅窗口内）+ 时长域闸 + 无除法 ｜ R5 ✓ 声明逐行同行双语注释
 *                         R6 ✓ 四态 ENUM + CASE + ELSE 兜底 ｜ R7 ✓ TON 实例 CASE 外无条件刷新
 * 修订历史 (Revision)   : 2026-11-23  v1.0.0  R77 首版（批次 B3 · 序号 12）
 * 验收向量 (Acceptance) : ① bGate=TRUE 时 fIn 由 10 变 20 → 当拍 fOut=20；
 *                         ② 随后 bGate=FALSE 且 fIn=99 → fOut 保持 20（不采纳）, bStale=FALSE（未超时）；
 *                         ③ bGate 持续 FALSE 超过 tMaxHold=T#1S → bStale=TRUE，fOut 仍保持 20；
 *                         ④ bGate=TRUE 且 fIn=NaN → uErrorId=16#0006_0002，bError=TRUE，fOut 冻结；
 *                         ⑤ tMaxHold=T#0S → bStale 恒 FALSE（显式屏蔽）。
 *==============================================================================*)

(*-----------------------------------------------------------------------------
 * 枚举: E_DL_GatedUpdState（门控更新状态机，归属 DL_Algo，与本件同文件，全库唯一属主）
 *-----------------------------------------------------------------------------
 * 过渡态说明：eInit --(首拍)--> eRun；eRun --(bGate=TRUE)--> eRun（更新）；
 * eRun --(bGate=FALSE)--> eRun（保持）；任一态 --(bEnable=FALSE)--> eHold；
 * 任一态 --(非有限/非法参数)--> eFault；eFault --(bEnable=FALSE 或 bReset)--> eInit。
 *----------------------------------------------------------------------------*)
TYPE E_DL_GatedUpdState :
(
    eInit  := 0,    // 首扫 / 复位后：输出直取输入 / First scan or after reset: output follows input
    eRun   := 10,   // 运行态：窗口内更新、窗口外保持 / Running: update inside window, hold outside
    eHold  := 20,   // 保持态：未使能，输出冻结 / Hold: disabled, output frozen
    eFault := 99    // 故障态：输出冻结，等待 bEnable 跌落或 bReset / Fault: frozen until cleared
);
END_TYPE

FUNCTION_BLOCK FB_DL_GatedUpdateFilter
VAR_INPUT
    bEnable  : BOOL := FALSE;      // 使能，FALSE 冻结输出 / Enable, FALSE freezes output
    bReset   : BOOL := FALSE;      // 复位到当前输入（单拍有效） / Reset to current input, single scan
    fIn      : LREAL := 0.0;       // 采样输入 [EU] / Sampling input [EU]
    bGate    : BOOL := FALSE;      // 窗口使能，TRUE = 本拍采纳输入 / Gate, TRUE adopts the input this scan
    tMaxHold : TIME := T#5S;       // 允许的最大保持时长，T#0S = 不判陈旧 [s] / Max hold duration, zero disables staleness
END_VAR
VAR_OUTPUT
    fOut         : LREAL;   // 门控输出 [EU] / Gated output [EU]
    bStale       : BOOL;    // 数据陈旧标志（信息级） [-] / Data staleness flag, info level
    tHeldElapsed : TIME;    // 已保持时长 [s] / Elapsed hold duration
    bValid       : BOOL;    // 输出有效标志 [-] / Output valid flag
    bError       : BOOL;    // 故障标志，与 uErrorId 联动 [-] / Fault flag coupled with uErrorId
    uErrorId     : UDINT;   // 故障码，0 = 无故障 [-] / Error code, zero means healthy
END_VAR
VAR
    tonHold  : TON;                  // 保持时长计时器（无条件每周期刷新） / Hold timer, refreshed unconditionally
    eState   : E_DL_GatedUpdState;   // 状态机当前状态 [-] / Current state
END_VAR
VAR CONSTANT
    DL_GUF_ZERO_L : LREAL := 0.0;    // 零基准（含非有限判零） [-] / Zero base including non-finite probe
    DL_GUF_ZERO_T : TIME := T#0S;    // 时长零基准 [s] / Zero duration base
END_VAR

(* —— 段 1：时长域闸（不中断扫描，只钳位并置信息码） —— *)
uErrorId := 16#0006_0000;                          // 预置无故障 / Preset healthy
IF tMaxHold < DL_GUF_ZERO_T THEN
    tMaxHold := DL_GUF_ZERO_T;                     // 负时长钳到零 / Negative duration clamped
    uErrorId := 16#0006_0001;                      // 信息级：时长已钳位 / Info: duration clamped
END_IF

(* —— 段 2：非有限防御（仅窗口内读取 fIn；窗口外输入无意义，不判故障） —— *)
IF bEnable AND bGate THEN
    IF (fIn <> fIn) OR ((fIn - fIn) <> DL_GUF_ZERO_L) THEN
        eState   := eFault;                        // 强制故障态 / Force fault state
        uErrorId := 16#0006_0002;                  // 故障级：窗口内输入非有限 / Fault: non-finite input inside window
    END_IF
END_IF

(* —— 段 3：复位请求 → 回首扫 —— *)
IF bReset THEN
    eState := eInit;
END_IF

(* —— 段 4：状态派生 —— *)
IF NOT bEnable THEN
    eState := eHold;                               // 未使能：冻结 / Disabled: freeze
ELSIF eState = eFault THEN
    eState := eFault;                              // 故障态保持 / Fault holds
ELSIF eState = eInit THEN
    eState := eInit;                               // 首扫保持一拍 / Init holds one scan
ELSE
    eState := eRun;
END_IF

(* —— 段 5：计时器无条件每周期刷新（R7 硬要求，位于 CASE 之外） —— *)
(* 计时条件：已使能、非故障、且当前不在窗口内（窗口外才累计「陈旧」时长） *)
(* Timer runs only when enabled, healthy, and outside the gate window *)
tonHold(IN := bEnable AND (eState <> eFault) AND (NOT bGate), PT := tMaxHold);

(* —— 段 6：主状态机（CASE 覆盖 + ELSE 兜底） —— *)
CASE eState OF

    eInit:
        fOut         := fIn;                       // 首拍直取输入 / First scan follows input
        bStale       := FALSE;                     // 首拍不判陈旧 / No staleness on first scan
        tHeldElapsed := tonHold.ET;
        bValid       := TRUE;
        eState       := eRun;

    eRun:
        IF bGate THEN
            fOut   := fIn;                         // 窗口内：原样采纳（无失真、无滞后） / Inside window: adopt raw
            bStale := FALSE;                       // 数据新鲜 / Data fresh
        ELSE
            (* 窗口外：fOut 保持上拍值，不做任何改写（保持语义核心） *)
            (* Outside window: hold previous output unchanged, core hold semantics *)
            IF (tMaxHold = DL_GUF_ZERO_T) THEN
                bStale := FALSE;                   // T#0S = 不判陈旧（显式屏蔽） / Zero disables staleness
            ELSE
                bStale := tonHold.Q;               // 超时才置陈旧 / Stale only after timeout
            END_IF
        END_IF
        tHeldElapsed := tonHold.ET;
        bValid       := TRUE;

    eHold:
        (* 未使能：输出与计时保持冻结 / Disabled: output and timer frozen *)
        bStale       := bStale;
        tHeldElapsed := tonHold.ET;
        bValid       := FALSE;

    eFault:
        (* 故障态：输出冻结保持上拍值（不推 0），计时器仍刷新 / Fault: output frozen, timer refreshed *)
        tHeldElapsed := tonHold.ET;
        bValid       := FALSE;

    ELSE
        eState   := eFault;
        bValid   := FALSE;
        uErrorId := 16#0006_0005;                  // 故障级：非法状态 / Fault: illegal state

END_CASE;

(* —— 段 7：出口映射（bError 与 uErrorId 同源；bStale 为信息级不置 bError） —— *)
bError := (uErrorId <> 16#0006_0000) AND (uErrorId <> 16#0006_0001);

END_FUNCTION_BLOCK

(* ---- FB_DL_HashBucketIndex.st ---- *)
(* ===========================================================================
   组件名   : FB_DL_HashBucketIndex
   分类     : DL_Algo / 哈希桶索引映射
   一句话   : 把 32 位哈希映射到桶号，支持掩码模式并要求桶数为 2 的幂，桶数为 0 时拒绝
   复杂度   : 2        版本 : v1.0.0        日期 : 2026-11-24
   开源溯源 : 无（clean-room 自研，未借鉴任何开源实现）
   输入契约 : dwHash 32 位哈希值；iBucketCount 桶数 1..32767；xUseMask TRUE=掩码模式
   输出契约 : iBucket 桶号 0..iBucketCount−1；dwMask 生效掩码（掩码模式）
              xMaskMode 实际使用掩码；xValid 输入有效
              iErrorCode 0=正常 1=桶数非正 2=掩码模式下桶数非 2 的幂
   修改记录 : v1.0.0 2026-11-24 初版
   =========================================================================== *)

FUNCTION_BLOCK FB_DL_HashBucketIndex
VAR_INPUT
    dwHash : DWORD := 0;               // 32 位哈希值 | 32 bit hash value
    iBucketCount : INT := 16;          // 桶数 1..32767 | bucket count 1..32767
    xUseMask : BOOL := TRUE;           // TRUE=掩码模式 | TRUE=mask mode
END_VAR
VAR_OUTPUT
    iBucket : INT;                     // 映射得到的桶号 | mapped bucket index
    dwMask : DWORD;                    // 生效掩码 | effective mask
    xMaskMode : BOOL;                  // 是否实际使用掩码 | mask actually used
    xValid : BOOL;                     // 输入有效标志 | inputs valid flag
    iErrorCode : INT;                  // 故障码 0=无故障 | error code
END_VAR
VAR
    dwCount : DWORD;                   // 桶数无符号形式 | bucket count as dword
    dwM : DWORD;                       // 候选掩码 | candidate mask
    dwBucket : DWORD;                  // 桶号工作值 | bucket working value
    _xPow2 : BOOL;                     // 桶数是否 2 的幂 | bucket count is power of two
END_VAR

// ---- 输出预置 ----
iBucket := 0;
dwMask := 0;
xMaskMode := FALSE;
xValid := FALSE;
iErrorCode := 0;

// ---- 桶数为 0 保护：直接拒绝，禁止进入任何除法/取模 ----
IF iBucketCount <= 0 THEN
    iErrorCode := 1;
ELSE
    dwCount := INT_TO_DWORD(iBucketCount);

    // ---- 掩码模式：桶数必须是 2 的幂，否则掩码无意义 ----
    IF xUseMask THEN
        dwM := dwCount - 1;
        _xPow2 := ((dwCount AND dwM) = 0) AND (dwCount > 1);
        IF _xPow2 THEN
            dwMask := dwM;
            xMaskMode := TRUE;
            dwBucket := dwHash AND dwM;            // 掩码取低位
            xValid := TRUE;
        ELSE
            iErrorCode := 2;                       // 非 2 的幂，掩码模式不可用
        END_IF
    ELSE
        // ---- 取模模式：桶数已保证非零，UDINT 取模避免有符号溢出 ----
        dwBucket := UDINT_TO_DWORD(DWORD_TO_UDINT(dwHash) MOD DWORD_TO_UDINT(dwCount));
        xValid := TRUE;
    END_IF

    IF xValid THEN
        // ---- 结果钳位：防御性保证桶号落在 [0, 桶数−1] ----
        IF dwBucket >= dwCount THEN
            dwBucket := dwCount - 1;
        END_IF
        iBucket := DWORD_TO_INT(dwBucket);         // 已小于 32767，转换安全
    END_IF
END_IF
END_FUNCTION_BLOCK

(* ---- FB_DL_HeatExchangerCtrl.st ---- *)
// =====================================================================
// FB_DL_HeatExchangerCtrl.st
// 换热器出口温度分程控制（低温段蒸汽阀加热 / 高温段凝水阀冷却）
// Heat exchanger split-range outlet temperature control FB
// 码位: 16#0002_3724 ~ 16#0002_3728 (本件独占 5 槽)
// 修改记录: R29 初版 (按 DISPATCH_R29 序 6)
// =====================================================================
FUNCTION_BLOCK FB_DL_HeatExchangerCtrl
VAR_INPUT
    bEnable       : BOOL  := FALSE;    // 使能 / Enable
    bPvValid      : BOOL  := FALSE;    // 温度有效 / PV valid
    fPv_C         : REAL  := 20.0;     // 出口温度 -20~250 ℃ / Outlet temperature [degC]
    fSp_C         : REAL  := 80.0;     // 设定 0~200 ℃ / Setpoint [degC]
    fDeadBand_C   : REAL  := 1.0;      // 分程死区 0~10 K / Split dead band [K]
    fKp           : REAL  := 3.0;      // 比例增益 0.1~50 %/K / Gain [%/K]
    fTi_s         : REAL  := 60.0;     // 积分时间 >0 s / Integral time [s]
    fBiasPct      : REAL  := 2.0;      // 交接偏置 0~20 % / Handover bias [%]
    fCondSafe_pct : REAL  := 30.0;     // 凝水阀安全位 0~100 % / Condensate safe position [%]
    bSteamAvail   : BOOL  := TRUE;     // 蒸汽可用 / Steam available
    bCondAvail    : BOOL  := TRUE;     // 凝水可用 / Condensate available
    bReset        : BOOL  := FALSE;    // 故障复位（电平持有一个周期即生效）/ Fault reset, level held for one cycle
    tCycle        : TIME  := T#200MS;  // 周期 T#20MS~T#5S / Cycle [s]
END_VAR
VAR_OUTPUT
    fSteamOut_pct : REAL;               // 蒸汽阀 0~100 % / Steam valve [%]
    fCondOut_pct  : REAL;               // 凝水阀 0~100 % / Condensate valve [%]
    fErr_C        : REAL;               // 温度偏差 K / Deviation [K]
    bSplitActive  : BOOL;               // 分程动作中 / Split active
    bDegraded     : BOOL;               // 单支路降级 / Degraded single branch
    eErr          : UDINT;              // 错误码 / Error code
END_VAR
VAR
    fIntegral     : REAL  := 0.0;       // 积分项 / Integral term [%]
    fTerm         : REAL  := 0.0;       // 本支路计算项 / Branch computed term [%]
    fIncr         : REAL  := 0.0;       // 本拍积分增量 / Integral increment this cycle [%]
    tCycleS       : REAL;               // 周期秒值 / Cycle in seconds [s]
    fDbSafe       : REAL;               // 兜底死区 / Sanitized dead band [K]
    bMutexLatch   : BOOL  := FALSE;     // 分程互斥失效锁存 / Split mutex fault latch
    xFirstScan    : BOOL  := TRUE;      // 首扫标记 / First-scan flag
END_VAR

// ---------------------------------------------------------------------
// 代码位表（本件独占，勿复用）:
//   16#0002_3724 信息 正常运行
//   16#0002_3725 故障 输入非有限 / tCycle 非法 / fTi_s ≤ 0（含 PV=NaN 安全侧分支）
//   16#0002_3726 故障 fKp ≤ 0 / fDeadBand_C < 0 / fBiasPct < 0（组态错）
//   16#0002_3727 信息 单支路降级（蒸汽或凝水不可用）→ bDegraded=TRUE；bPvValid=FALSE 安全侧同登记
//   16#0002_3728 故障 双阀同时 >0.5 % 且 ABS(fErr_C) > fDeadBand_C → 双阀归 0 锁存，解除=bReset 且带内
// ---------------------------------------------------------------------

// ---- 周期转秒 / Cycle to seconds ----
tCycleS := TIME_TO_REAL(tCycle) / 1000.0;   // 秒值 / Seconds [s]

// ---- 非有限与时域合法性闸（故障级）/ Finite and time-domain gate ----
IF (tCycle = T#0MS) OR (tCycleS < 0.02) OR (tCycleS > 5.0)
   OR (fTi_s <= 0.0)
   OR (fPv_C <> fPv_C) OR (ABS(fPv_C) >= 1.0E12)
   OR (fSp_C <> fSp_C) OR (ABS(fSp_C) >= 1.0E12)
   OR (fCondSafe_pct <> fCondSafe_pct) OR (ABS(fCondSafe_pct) >= 1.0E12) THEN
    fSteamOut_pct := 0.0;       // 蒸汽阀安全关闭 / Steam safe closed
    fCondOut_pct  := fCondSafe_pct; // 凝水阀安全位 / Condensate safe position
    bSplitActive  := FALSE;     // 分程退出 / Split inactive
    bDegraded     := TRUE;      // 登记降级 / Mark degraded
    eErr          := 16#0002_3725;  // 故障码 / Fault code
    RETURN;                     // 本拍结束 / End of cycle
END_IF

// ---- 组态错闸 / Configuration fault gate ----
IF (fKp <= 0.0) OR (fDeadBand_C < 0.0) OR (fBiasPct < 0.0) THEN
    fSteamOut_pct := 0.0;       // 蒸汽阀关闭 / Steam closed
    fCondOut_pct  := 0.0;       // 凝水阀关闭 / Condensate closed
    bSplitActive  := FALSE;     // 分程退出 / Split inactive
    eErr          := 16#0002_3726;  // 故障码 / Fault code
    RETURN;                     // 本拍结束 / End of cycle
END_IF

// ---- 死区兜底：0 按 0.5 K 防抖振 / Dead-band fallback: 0 to 0.5 K ----
IF fDeadBand_C = 0.0 THEN
    fDbSafe := 0.5;             // 兜底 0.5 K / Fallback 0.5 K
ELSE
    fDbSafe := fDeadBand_C;     // 原值 / As-is
END_IF

// ---- 首扫初始化 / First-scan initialization ----
IF xFirstScan THEN
    fSteamOut_pct := 0.0;       // 蒸汽阀初始关 / Steam init closed
    fCondOut_pct  := 0.0;       // 凝水阀初始关 / Condensate init closed
    fIntegral     := 0.0;       // 积分清零 / Integral cleared
    xFirstScan    := FALSE;     // 清标记 / Clear flag
END_IF

// ---- 使能撤销：双阀回关 / Disable: both valves closed ----
IF NOT bEnable THEN
    fSteamOut_pct := 0.0;       // 蒸汽阀关 / Steam closed
    fCondOut_pct  := 0.0;       // 凝水阀关 / Condensate closed
    bSplitActive  := FALSE;     // 分程退出 / Split inactive
    bDegraded     := FALSE;     // 降级复位 / Reset degraded
    eErr          := 16#0002_3724;  // 信息级：空闲正常 / Info: idle normal
    RETURN;                     // 本拍结束 / End of cycle
END_IF

// ---- 偏差计算 / Deviation computation ----
fErr_C := fSp_C - fPv_C;        // 偏差 = SP - PV / Deviation [K]

// ---- 分程互斥失效锁存与解除 / Split mutex latch and release ----
IF bMutexLatch THEN
    // 锁存中：双阀归 0，解除 = bReset 且 ABS(fErr_C) ≤ fDbSafe / Latched: valves 0, release on reset+in-band
    fSteamOut_pct := 0.0;       // 蒸汽阀归 0 / Steam zero
    fCondOut_pct  := 0.0;       // 凝水阀归 0 / Condensate zero
    bSplitActive  := FALSE;     // 分程退出 / Split inactive
    eErr := 16#0002_3728;       // 故障码回放 / Fault code replay
    IF bReset AND (ABS(fErr_C) <= fDbSafe) THEN
        bMutexLatch := FALSE;   // 解除锁存 / Release latch
        fIntegral   := 0.0;     // 积分清零重新起步 / Clear integral
    END_IF
    RETURN;                     // 本拍结束 / End of cycle
END_IF

// ---- PV 无效安全侧：蒸汽关、凝水安全位 / PV invalid safe side ----
IF NOT bPvValid THEN
    fSteamOut_pct := 0.0;       // 蒸汽关 / Steam closed
    fCondOut_pct  := fCondSafe_pct; // 凝水安全位 / Condensate safe
    bSplitActive  := FALSE;     // 分程退出 / Split inactive
    bDegraded     := TRUE;      // 登记降级（信息级，不置故障）/ Mark degraded (info only)
    eErr          := 16#0002_3727;  // 信息级：降级 / Info: degraded
    RETURN;                     // 本拍结束 / End of cycle
END_IF

// ---- 单支路可用性降级登记 / Single-branch availability degrade ----
bDegraded := (NOT bSteamAvail) OR (NOT bCondAvail);  // 降级标志 / Degraded flag

// ---- 分程 PI 计算（内联，交接偏置防抢动）/ Split-range PI with handover bias ----
bSplitActive := FALSE;          // 默认分程未动作 / Default inactive
IF fErr_C > fDbSafe THEN
    // 低温段：开蒸汽阀加热 / Low side: steam heating
    fIncr := (fErr_C / fTi_s) * tCycleS;    // 积分增量 / Integral increment [%]
    // 抗饱和：蒸汽支路到 100 % 边沿停同向积分 / Anti-windup at 100 %
    IF (fSteamOut_pct >= 100.0) AND (fIncr > 0.0) THEN
        fIncr := 0.0;           // 停同向积分 / Freeze integral
    END_IF
    fIntegral := fIntegral + fIncr;     // 积分累计 / Integrate
    fTerm := fKp * (fErr_C - fDbSafe) + fIntegral + fBiasPct;   // 计算项含交接偏置 / Term with bias [%]
    IF fTerm < 0.0 THEN
        fTerm := 0.0;           // 下限钳 / Lower clamp
    ELSIF fTerm > 100.0 THEN
        fTerm := 100.0;         // 上限钳（下一拍抗饱和生效）/ Upper clamp
    END_IF
    IF bSteamAvail THEN
        fSteamOut_pct := fTerm; // 蒸汽阀输出 / Steam output
    ELSE
        fSteamOut_pct := 0.0;   // 蒸汽不可用 → 支路 0 / Steam unavailable
    END_IF
    fCondOut_pct := 0.0;        // 凝水阀关 / Condensate closed
    bSplitActive := TRUE;       // 分程动作中 / Split active
    eErr := 16#0002_3724;       // 信息级：正常 / Info: normal
ELSIF fErr_C < -fDbSafe THEN
    // 高温段：开凝水阀冷却 / High side: condensate cooling
    fIncr := (-fErr_C / fTi_s) * tCycleS;   // 积分增量 / Integral increment [%]
    // 抗饱和：凝水支路到 100 % 边沿停同向积分 / Anti-windup at 100 %
    IF (fCondOut_pct >= 100.0) AND (fIncr > 0.0) THEN
        fIncr := 0.0;           // 停同向积分 / Freeze integral
    END_IF
    fIntegral := fIntegral + fIncr;     // 积分累计 / Integrate
    fTerm := fKp * (-fErr_C - fDbSafe) + fIntegral + fBiasPct;  // 计算项含交接偏置 / Term with bias [%]
    IF fTerm < 0.0 THEN
        fTerm := 0.0;           // 下限钳 / Lower clamp
    ELSIF fTerm > 100.0 THEN
        fTerm := 100.0;         // 上限钳 / Upper clamp
    END_IF
    IF bCondAvail THEN
        fCondOut_pct := fTerm;  // 凝水阀输出 / Condensate output
    ELSE
        fCondOut_pct := 0.0;    // 凝水不可用 → 支路 0 / Condensate unavailable
    END_IF
    fSteamOut_pct := 0.0;       // 蒸汽阀关 / Steam closed
    bSplitActive := TRUE;       // 分程动作中 / Split active
    eErr := 16#0002_3724;       // 信息级：正常 / Info: normal
ELSE
    // 死区带内：双阀同关 / In dead band: both closed
    fSteamOut_pct := 0.0;       // 蒸汽阀关 / Steam closed
    fCondOut_pct  := 0.0;       // 凝水阀关 / Condensate closed
    eErr := 16#0002_3724;       // 信息级：正常 / Info: normal
END_IF

// ---- 分程互斥闸（防御性复核，越过分程死区双阀非零 → 故障锁存）/ Mutex recheck ----
IF (fSteamOut_pct > 0.5) AND (fCondOut_pct > 0.5) AND (ABS(fErr_C) > fDbSafe) THEN
    fSteamOut_pct := 0.0;       // 双阀归 0 / Both valves zero
    fCondOut_pct  := 0.0;       // 双阀归 0 / Both valves zero
    bMutexLatch   := TRUE;      // 锁存 / Latch
    eErr          := 16#0002_3728;  // 故障码 / Fault code
END_IF

// ---- 单支路降级信息级覆盖 / Degraded info code override ----
IF bDegraded AND (eErr = 16#0002_3724) THEN
    eErr := 16#0002_3727;       // 信息级：单支路降级 / Info: degraded
END_IF

END_FUNCTION_BLOCK

(* ---- FB_DL_HighPassFilter.st ---- *)
(*==============================================================================
 * 组件名称 (Component)  : FB_DL_HighPassFilter
 * 所属子库 (Sublibrary) : DL_Algo
 * 当前版本 (Version)    : 1.0.0
 * 兼容性   (Platform)   : CODESYS 3.5 / TwinCAT 3 / 汇川 InoProShop / Machine Expert
 *                         仅依赖 Standard.library（MIN / MAX / ABS / LIMIT），
 *                         零厂商方言
 * 功能描述 (Function)   : 一阶高通数字滤波器（HP1）。递推式
 *                         fOut := fAlpha * (fOutPrev + fIn - fInPrev)，
 *                         其中 fAlpha := tTf / (tTf + fDt)。剥离静态偏置、
 *                         提取动态分量：振动 / 位移传感器趋势分量剥离、
 *                         皮带秤动态分量提取、结露监测的缓变漂移滤除。
 *                         含输出限幅（rOutMin/rOutMax 对调防御）、
 *                         tTimeConst=0 全通差分、首扫防上电脉冲、
 *                         bTrack 跟踪时输出清零并同步历史。
 * 开源溯源 (Origin)     : 原创实现。算法思想源自 LGF HP1 与一阶高通差分
 *                         教科书推导（clean-room），按本库故障码体系重写。
 * 设计验证 (Verified)   : tTf=0.1s、fDt=0.01s：fAlpha=0.909091；
 *                         正弦 1Hz 输入稳态增益约 0.532018（python 核验）；
 *                         直流阶跃 0->5.0 输入：第 1 拍动态分量 4.545455，
 *                         第 50 拍衰减至 0.042593（静态偏置被隔离并归零）。
 * 验收向量 (Acceptance) :
 *   V1 fAlpha=0.909091（tTf=0.1s fDt=0.01s，容差 1E-4）
 *   V2 直流阶跃 0->5.0：50 拍后 fOut < 0.5（动态分量快速归零）
 *   V3 tTimeConst=T#0S：fOut=fIn-fInPrev（全通差分）
 *   V4 bTrack=TRUE：当拍 fOut=0.0 且历史同步，回自动无脉冲
 *   V5 输出 12.0 超 rOutMax=10.0：当拍钳位 10.0，uErrorId=16#0002_0001
 *   V6 fIn 非有限值：拒绝更新并复位历史，uErrorId=16#0002_0004
 * 本文件内含       : TYPE  E_DL_HpfState（配套枚举，归属 DL_Algo）
 *                    FB    FB_DL_HighPassFilter
 * 依赖     (Depends)    : 无 DL_ 内部依赖；Standard.library 数学算符
 * 红线自检 (Redline)    : R1 ✓ 零全局变量表与外部变量引用 ｜ R2 ✓ 零物理 IO 地址直写
 *                         R3 ✓ 纯 IEC 61131-3 ｜ R4 ✓ 钳位+容差+非有限值拒绝+对调防御
 *                         R5 ✓ 全变量中英双语同行注释 ｜ R6 ✓ 四态 ENUM+CASE+ELSE
 *                         R7 N/A（无定时器与边沿检测实例）
 * 修订历史 (Revision)   :
 *   2026-11-15  v1.0.0  首版入库（Round 04 · Phase 3 · DL_Algo 批次）
 *============================================================================*)

(*-----------------------------------------------------------------------------
 * 枚举: E_DL_HpfState（归属 DL_Algo，与 FB_DL_HighPassFilter 同文件）
 * 含义: 高通滤波状态机离散状态。纯线性滤波采用「状态派生 + CASE 覆盖 + ELSE」
 *       结构：状态由使能 / 跟踪 / 首扫信号派生，CASE 保证每态行为显式可审计。
 *----------------------------------------------------------------------------*)
TYPE E_DL_HpfState :
(
    eInit  := 0,    // 首扫态：输出清零并同步输入历史，防上电脉冲 / First scan: output zeroed with input history synced, no power-up pulse
    eRun   := 10,   // 运行态：按 fAlpha 递推提取动态分量 / Running: recursive dynamic component extraction with fAlpha
    eTrack := 20,   // 跟踪态：输出清零并同步历史，投切无脉冲 / Tracking: output zeroed with history synced, bumpless transfer
    eFault := 99    // 故障兜底态：非法状态进入，输出安全值并置故障码 / Fault fallback: entered from illegal states, safe output plus error code
);
END_TYPE

(*==============================================================================
 * 功能块: FB_DL_HighPassFilter
 * 调用约定: 每个采样周期无条件调用一次；tSampleTime 由调用方显式给定，
 *           严禁依赖隐式扫描周期做差分递推；多实例可并行互不干扰。
 * 滞后披露: 截止频率 fc = 1/(2*pi*tTf)；低于 fc 的缓变分量被衰减，
 *           时间常数越大截止频率越低、保留的低频动态越丰富。
 * 限幅披露: 输出限幅为工程防护（防差分尖峰打穿下游量程），非滤波语义；
 *           rOutMin > rOutMax 时二者对调并置公共钳位码，不中断扫描。
 *============================================================================*)
FUNCTION_BLOCK FB_DL_HighPassFilter
VAR_INPUT
    bEnable     : BOOL := FALSE;      // 使能，FALSE 时输出置 0 / Enable, FALSE forces output to zero
    fIn         : REAL := 0.0;        // 原始采样输入 [EU] / Raw sampling input [EU]
    tTimeConst  : TIME := T#1S;       // 高通时间常数 [s]，越大截止频率越低；T#0S=全通差分 / High-pass time constant [s], larger means lower cutoff; T#0S = all-pass difference
    tSampleTime : TIME := T#100MS;    // 采样周期，小于 10ms 钳位 / Sampling period, clamped to 10ms minimum
    rOutMin     : REAL := -1.0E10;    // 输出下限 [EU] / Output lower limit [EU]
    rOutMax     : REAL := 1.0E10;     // 输出上限 [EU] / Output upper limit [EU]
    bTrack      : BOOL := FALSE;      // 跟踪使能，TRUE 时输出清零并同步历史 / Track enable, TRUE zeroes output and synchronizes history
    fTrackValue : REAL := 0.0;        // 跟踪目标值 [EU]，跟踪语义为清零基线 / Track target value [EU], tracking zeroes the baseline
END_VAR
VAR_OUTPUT
    fOut        : REAL;               // 动态分量输出 [EU] / Dynamic component output [EU]
    fAlpha      : REAL;               // 当前滤波系数 [0..1]，诊断用 / Current filter coefficient [0..1], diagnostic
    bValid      : BOOL;               // 输出有效标志，首扫未完成时为 FALSE / Output valid flag, FALSE before first scan completes
    bError      : BOOL;               // 故障标志，与 uErrorId 联动 / Fault flag, coupled with uErrorId
    uErrorId    : UDINT;              // 故障码，0 = 无故障 / Error code, 0 = no error
END_VAR
VAR
    fInPrev     : REAL := 0.0;        // 上拍输入历史 [EU]，首扫同步防尖峰 / Previous input history [EU], synced at first scan
    fTfEff      : REAL;               // 钳位后的生效时间常数 [s] / Effective clamped time constant [s]
    fDt         : REAL;               // 采样周期秒值 [s] / Sampling period in seconds [s]
    fTfRaw      : REAL;               // 时间常数换算秒值（钳位前）[s] / Time constant in seconds before clamping [s]
    fOutLo      : REAL;               // 排序后的输出下限 [EU] / Ordered output lower limit [EU]
    fOutHi      : REAL;               // 排序后的输出上限 [EU] / Ordered output upper limit [EU]
    eState      : E_DL_HpfState;      // 状态机当前状态 / Current state of the state machine
END_VAR
VAR CONSTANT
    DL_HPF_TF_MAX  : REAL := 3600.0;  // 时间常数上限 [s]，超限钳位防过度迟滞 / Time constant upper clamp [s], prevents excessive lag
    DL_HPF_DT_MIN  : REAL := 0.01;    // 采样周期防御下限 [s] / Defensive sampling period lower bound [s]
    DL_HPF_INF_MAX : REAL := 1.0E30;  // 有限值判定幅值上限 [EU] / Magnitude bound for finite-value check [EU]
END_VAR

(*------------------------------------------------------------------------------
 * 段 1｜参数钳位（不中断扫描）：周期下限 / 时间常数域 / 限幅对调
 *      Parameter clamping without scan interruption: period floor, constant range, limit swap
 *-----------------------------------------------------------------------------*)
uErrorId := 16#0002_0000;

IF tSampleTime < T#10MS THEN
    fDt      := DL_HPF_DT_MIN;                       // 周期过小钳位到 10ms / Too small period clamped to 10ms
    uErrorId := 16#0002_0002;                        // 采样周期非法已钳位 / Invalid sampling period clamped
ELSE
    fDt := TIME_TO_REAL(tSampleTime) / 1000.0;       // TIME 换算秒值 / Convert TIME to seconds
END_IF

fTfRaw := TIME_TO_REAL(tTimeConst) / 1000.0;         // 时间常数换算秒值 / Convert time constant to seconds

IF (fTfRaw < 0.0) OR (fTfRaw > DL_HPF_TF_MAX) THEN
    fTfEff   := MIN(MAX(fTfRaw, 0.0), DL_HPF_TF_MAX); // 双侧钳位到合法域 / Two-sided clamp into valid range
    uErrorId := 16#0002_1201;                        // 时间常数非法已钳位 / Invalid time constant clamped
ELSE
    fTfEff := fTfRaw;                                // 合法参数原值生效 / Valid parameter applied as-is
END_IF

(* 限幅上下限对调防御：传反不中断扫描，排序后生效并置公共钳位码 *)
(* Limit swap defense: reversed limits are reordered without scan interruption *)
IF rOutMin > rOutMax THEN
    fOutLo   := rOutMax;
    fOutHi   := rOutMin;
    uErrorId := 16#0002_0001;                        // 参数越界已钳位（限幅对调） / Parameter out of range, limits swapped
ELSE
    fOutLo := rOutMin;
    fOutHi := rOutMax;
END_IF

(*------------------------------------------------------------------------------
 * 段 2｜滤波系数计算（防除零）：fAlpha = fTf/(fTf+fDt)
 *      Filter coefficient with divide-by-zero guard: fAlpha = fTf/(fTf+fDt)
 *      tTimeConst=0 时 fAlpha=0，全通差分语义与 V3 向量对应
 *-----------------------------------------------------------------------------*)
IF fTfEff <= 1.0E-6 THEN
    fAlpha := 0.0;                                   // 零时间常数：全通差分系数 / Zero constant: all-pass difference coefficient
ELSE
    fAlpha := MIN(MAX(fTfEff / (fTfEff + fDt), 0.0), 1.0); // 系数显式约束在 0 与 1 之间 / Coefficient constrained into 0..1
END_IF

(*------------------------------------------------------------------------------
 * 段 3｜非有限值防御：拒绝本拍更新、复位历史防差分尖峰（公共故障码）
 *      Non-finite defense: reject this cycle and reset history against spikes
 *-----------------------------------------------------------------------------*)
IF (fIn <> fIn) OR (ABS(fIn) > DL_HPF_INF_MAX) THEN
    uErrorId := 16#0002_0004;                        // 输入非有限值已拒绝 / Non-finite input rejected
    fInPrev  := 0.0;                                 // 历史复位，恢复后按首扫口径重建 / History reset, rebuilt like first scan after recovery
    bValid   := FALSE;
    bError   := TRUE;
    RETURN;
END_IF

(*------------------------------------------------------------------------------
 * 段 4｜主状态机（红线 R6）：状态派生 + CASE 覆盖 + ELSE 兜底
 *      Main state machine: state derived from signals, CASE covered with ELSE
 *-----------------------------------------------------------------------------*)
IF bTrack THEN
    eState := eTrack;                                // 跟踪请求优先级最高 / Track request has highest priority
ELSIF eState = eInit THEN
    eState := eInit;                                 // 首扫态保持，不被运行派生覆盖 / First scan state preserved from override
ELSIF eState = eFault THEN
    IF NOT bEnable THEN
        eState := eInit;                             // 使能跌落提供故障恢复路径 / Disabled input provides fault recovery path
    ELSE
        eState := eFault;                            // 故障态保持直至调用方处置 / Fault state holds until caller intervenes
    END_IF
ELSE
    eState := eRun;                                  // 常规运行态派生 / Normal running state derived
END_IF

CASE eState OF

    eInit:
        (* 首扫防上电脉冲：输出清零、输入历史与当前输入同步，差分基差为零 *)
        (* First scan power-up pulse guard: output zeroed, history synced to current input *)
        fOut    := 0.0;
        fInPrev := fIn;
        bValid  := FALSE;                            // 首扫未完成，输出尚不可信 / First scan unfinished, output not trustworthy yet
        eState  := eRun;                             // 下一拍进入运行态 / Move to running state next cycle

    eTrack:
        (* 无扰跟踪：输出清零、历史同步，回自动时差分基差为零无脉冲 *)
        (* Bumpless tracking: output zeroed, history synced, no pulse on resume *)
        fOut    := 0.0;
        fInPrev := fIn;
        bValid  := TRUE;
        eState  := eRun;

    eRun:
        IF NOT bEnable THEN
            (* 使能失效语义：输出置 0，历史同步防止恢复使能时残留脉冲 *)
            (* Disabled semantics: output zeroed, history synced to avoid resume pulses *)
            fOut    := 0.0;
            fInPrev := fIn;
            bValid  := FALSE;
        ELSE
            IF fAlpha <= 1.0E-6 THEN
                (* 全通差分：tTimeConst=0，输出为当拍与上拍之差 *)
                (* All-pass difference: zero time constant, output is cycle-to-cycle difference *)
                fOut := fIn - fInPrev;
            ELSE
                (* 一阶高通递推：fOut := fAlpha*(fOutPrev + fIn - fInPrev) *)
                (* First-order high-pass recursion per specification formula *)
                fOut := fAlpha * (fOut + fIn - fInPrev);
            END_IF

            (* 输出限幅：双侧钳位防差分尖峰打穿下游量程 *)
            (* Output limiting: two-sided clamp against downstream range breakthrough *)
            fOut := LIMIT(fOutLo, fOut, fOutHi);

            fInPrev := fIn;                          // 输入历史右移一位 / Shift input history by one
            bValid  := TRUE;
        END_IF

    eFault:
        (* 故障兜底：输出保持安全值 0，等待调用方修正后经使能跌落恢复 *)
        (* Fault fallback: output holds safe value 0, recovers via disabled input *)
        fOut   := 0.0;
        bValid := FALSE;

    ELSE
        (* 非法状态拦截：任何未定义枚举值一律进故障态并置公共兜底码 *)
        (* Illegal state interception: undefined enum values go to fault with code *)
        eState   := eFault;
        fOut     := 0.0;
        bValid   := FALSE;
        uErrorId := 16#0002_0005;

END_CASE;

(* 故障标志统一出口：与故障码严格联动，0 即无故障 *)
(* Unified fault flag outlet: strictly coupled with error code, zero means healthy *)
bError := (uErrorId <> 16#0002_0000);
END_FUNCTION_BLOCK

(* ---- FB_DL_HoldLastGoodFilter.st ---- *)
(*==============================================================================
 * 组件名称 (Component)  : FB_DL_HoldLastGoodFilter
 * 所属子库 (Sublibrary) : DL_Algo
 * 当前版本 (Version)    : 1.0.0
 * 兼容性   (Platform)   : CODESYS 3.5+ / TwinCAT 3 / 汇川 InoProShop / 施耐德 Machine Expert
 *                         仅依赖 Standard.library（TON），零厂商私有库
 * 功能描述 (Function)   : 坏值保持滤波（hold last good）。上游给出质量判据 bGood
 *                         （传感器在线 / 通信正常 / 量程内 / 非冻结），本件在判据有效时
 *                         采纳输入，判据失效时**输出上一有效值并累计失效时长**。
 *                         失效时长超过 tMaxBad 置 bTimedOut=TRUE（信息级，供上游降级决策），
 *                         输出**仍然保持**（不自动回落 0，避免下游把保持值当成真实 0）。
 *                         与 FB_DL_GatedUpdateFilter 的差别：那件按时间窗门控，
 *                         本件按数据质量门控；两者可串联（先门控再质量保持）。
 * 接口     (Interface)  : 输入 bEnable 使能、bReset 清「已获得首个有效值」标志、
 *                         fIn 采样输入 [EU]、bGood 质量判据（TRUE = 本拍可信）、
 *                         tMaxBad 允许的最大坏值持续时长 [s]；
 *                         输出 fOut 输出值 [EU]、bHolding 是否处于坏值保持、
 *                         bTimedOut 坏值超时（信息级）、tBadElapsed 已保持时长 [s]、
 *                         bValid 输出是否有可信值（从未得到过有效值时为 FALSE）、
 *                         bError 故障标志、uErrorId 故障码。
 * 边界     (Boundary)   : ① 属主边界：只做质量门控与保持，不判断质量本身
 *                         （bGood 由上游传感器诊断 / 量程判定给出，本件不越权推断）。
 *                         ② **从未得到过有效值**（bGood 从未 TRUE）时 bValid=FALSE 且 fOut=0，
 *                         这是唯一把输出置 0 的情形，已在头注释显式声明（名实双出口）。
 *                         ③ 非有限防御：仅当 bGood=TRUE 时读取 fIn；此时非有限 → 故障态
 *                         16#0007_0002（判据与数值矛盾，属上游逻辑错误，必须报）。
 *                         ④ tMaxBad < 0 钳到 T#0S 并置信息码 16#0007_0001；T#0S = 不判超时。
 *                         ⑤ **TON 无条件每周期调用**（R7），位于 CASE 之外。
 *                         ⑥ 零全局耦合（无 GVL / VAR_EXTERNAL / 物理地址）。
 * 分工声明 (Scope)      : 与 `FB_DL_GatedUpdateFilter` 分工：时间窗门控归那件、
 *                         质量门控归本件；与 `FB_DL_AnalogInputRedundancySel`（另批）分工：
 *                         双路择优归那件，本件不比较两路。
 * 来源标签 (Source Tag) : 原创实现（无外部代码引入）
 * 码表     (Codes)      : 16#0007_0000 无故障 / 16#0007_0001 坏值时长非法已钳位（信息级）/
 *                         16#0007_0002 判据有效但数值非有限（故障级）/ 16#0007_0005 非法状态（故障级）。
 * 红线自检 (Redline)    : R1 ✓ 零 GVL/VAR_EXTERNAL ｜ R2 ✓ 零 %I/%Q/%M ｜ R3 ✓ 纯 IEC 61131-3
 *                         R4 ✓ 非有限拒绝 + 时长域闸 + 无除法 ｜ R5 ✓ 声明逐行同行双语注释
 *                         R6 ✓ 四态 ENUM + CASE + ELSE 兜底 ｜ R7 ✓ TON 实例 CASE 外无条件刷新
 * 修订历史 (Revision)   : 2026-11-23  v1.0.0  R77 首版（批次 B3 · 序号 13）
 * 验收向量 (Acceptance) : ① bGood=TRUE, fIn=42.5 → fOut=42.5, bHolding=FALSE, bValid=TRUE；
 *                         ② 随后 bGood=FALSE, fIn=0.0 → fOut 保持 42.5, bHolding=TRUE, bValid=TRUE；
 *                         ③ bGood 持续 FALSE 超过 tMaxBad=T#2S → bTimedOut=TRUE，fOut 仍 42.5；
 *                         ④ 上电起 bGood 一直 FALSE → fOut=0.0, bValid=FALSE, bTimedOut 视时长；
 *                         ⑤ bGood=TRUE 且 fIn=NaN → uErrorId=16#0007_0002，bError=TRUE，fOut 冻结。
 *==============================================================================*)

(*-----------------------------------------------------------------------------
 * 枚举: E_DL_HoldGoodState（坏值保持状态机，归属 DL_Algo，与本件同文件，全库唯一属主）
 *----------------------------------------------------------------------------*)
TYPE E_DL_HoldGoodState :
(
    eInit  := 0,    // 首扫 / 复位后：尚未获得有效值 / First scan or after reset: no valid value yet
    eRun   := 10,   // 运行态：判据有效则采纳、失效则保持 / Running: adopt when good, hold when bad
    eHold  := 20,   // 保持态：未使能，输出冻结 / Hold: disabled, output frozen
    eFault := 99    // 故障态：输出冻结，等待 bEnable 跌落或 bReset / Fault: frozen until cleared
);
END_TYPE

FUNCTION_BLOCK FB_DL_HoldLastGoodFilter
VAR_INPUT
    bEnable : BOOL := FALSE;      // 使能，FALSE 冻结输出 / Enable, FALSE freezes output
    bReset  : BOOL := FALSE;      // 复位「已获有效值」标志（单拍有效） / Reset the valid-acquired flag, single scan
    fIn     : LREAL := 0.0;       // 采样输入 [EU] / Sampling input [EU]
    bGood   : BOOL := FALSE;      // 质量判据，TRUE = 本拍输入可信 / Quality flag, TRUE means trustworthy
    tMaxBad : TIME := T#5S;       // 允许的最大坏值持续时长，T#0S = 不判超时 [s] / Max bad duration, zero disables
END_VAR
VAR_OUTPUT
    fOut        : LREAL;   // 输出值（坏值期间保持） [EU] / Output value, held while bad
    bHolding    : BOOL;    // 是否处于坏值保持 [-] / Whether holding a previous value
    bTimedOut   : BOOL;    // 坏值超时（信息级） [-] / Bad-value timeout, info level
    tBadElapsed : TIME;    // 已保持时长 [s] / Elapsed hold duration
    bValid      : BOOL;    // 输出是否有可信值 [-] / Whether the output holds a trustworthy value
    bError      : BOOL;    // 故障标志，与 uErrorId 联动 [-] / Fault flag coupled with uErrorId
    uErrorId    : UDINT;   // 故障码，0 = 无故障 [-] / Error code, zero means healthy
END_VAR
VAR
    tonBad    : TON;                  // 坏值时长计时器（无条件每周期刷新） / Bad duration timer, refreshed unconditionally
    _bHasGood : BOOL;                 // 是否已获得过有效值 [-] / Whether a good value was ever acquired
    _fLastGood: LREAL;                // 上一有效值 [EU] / Last good value
    eState    : E_DL_HoldGoodState;   // 状态机当前状态 [-] / Current state
END_VAR
VAR CONSTANT
    DL_HGF_ZERO_L : LREAL := 0.0;    // 零基准（含非有限判零） [-] / Zero base including non-finite probe
    DL_HGF_ZERO_T : TIME := T#0S;    // 时长零基准 [s] / Zero duration base
END_VAR

(* —— 段 1：时长域闸（不中断扫描，只钳位并置信息码） —— *)
uErrorId := 16#0007_0000;                          // 预置无故障 / Preset healthy
IF tMaxBad < DL_HGF_ZERO_T THEN
    tMaxBad := DL_HGF_ZERO_T;                      // 负时长钳到零 / Negative duration clamped
    uErrorId := 16#0007_0001;                      // 信息级：时长已钳位 / Info: duration clamped
END_IF

(* —— 段 2：非有限防御（仅判据有效时读取 fIn；判据失效时输入无意义） —— *)
IF bEnable AND bGood THEN
    IF (fIn <> fIn) OR ((fIn - fIn) <> DL_HGF_ZERO_L) THEN
        eState   := eFault;                        // 判据与数值矛盾：报故障 / Contradiction between flag and value
        uErrorId := 16#0007_0002;                  // 故障级：判据有效但数值非有限 / Fault: good flag with non-finite value
    END_IF
END_IF

(* —— 段 3：复位请求 → 回首扫并清「已获有效值」标志 —— *)
IF bReset THEN
    eState    := eInit;
    _bHasGood := FALSE;                            // 清标志：需重新获得有效值 / Clear flag, must re-acquire
END_IF

(* —— 段 4：状态派生 —— *)
IF NOT bEnable THEN
    eState := eHold;                               // 未使能：冻结 / Disabled: freeze
ELSIF eState = eFault THEN
    eState := eFault;                              // 故障态保持 / Fault holds
ELSIF eState = eInit THEN
    eState := eInit;                               // 首扫保持一拍 / Init holds one scan
ELSE
    eState := eRun;
END_IF

(* —— 段 5：计时器无条件每周期刷新（R7 硬要求，位于 CASE 之外） —— *)
(* 计时条件：已使能、非故障、且当前判据失效（bad） *)
(* Timer runs only when enabled, healthy, and the quality flag is false *)
tonBad(IN := bEnable AND (eState <> eFault) AND (NOT bGood), PT := tMaxBad);

(* —— 段 6：主状态机（CASE 覆盖 + ELSE 兜底） —— *)
CASE eState OF

    eInit:
        IF bGood THEN
            _fLastGood := fIn;                     // 首个有效值 / First good value
            _bHasGood  := TRUE;
            fOut       := fIn;
            bHolding   := FALSE;
            bValid     := TRUE;
            eState     := eRun;                    // 已获有效值，进入运行态 / Enter running
        ELSE
            fOut     := DL_HGF_ZERO_L;             // 从未获得有效值：唯一置 0 的情形 / Only case that zeroes output
            bHolding := FALSE;
            bValid   := FALSE;                     // 明确声明：无可信值 / Explicitly no trustworthy value
            eState   := eRun;
        END_IF
        tBadElapsed := tonBad.ET;
        bTimedOut   := FALSE;

    eRun:
        IF bGood THEN
            _fLastGood := fIn;                     // 刷新上一有效值 / Refresh last good value
            _bHasGood  := TRUE;
            fOut       := fIn;                     // 采纳本拍输入 / Adopt current input
            bHolding   := FALSE;
            bValid     := TRUE;
            bTimedOut  := FALSE;                   // 判据恢复：超时标志清除（可达解除路径） / Timeout cleared
        ELSE
            fOut     := _fLastGood;                // 保持上一有效值 / Hold last good value
            bHolding := TRUE;
            bValid   := _bHasGood;                 // 无有效值历史时仍不可信 / Untrustworthy without history
            IF tMaxBad = DL_HGF_ZERO_T THEN
                bTimedOut := FALSE;                // T#0S = 不判超时 / Zero disables timeout
            ELSE
                bTimedOut := tonBad.Q;             // 超时才置位 / Set only after timeout
            END_IF
        END_IF
        tBadElapsed := tonBad.ET;

    eHold:
        (* 未使能：输出、保持标志与计时全部冻结 / Disabled: output, flags and timer all frozen *)
        tBadElapsed := tonBad.ET;
        bValid      := FALSE;

    eFault:
        (* 故障态：输出冻结保持上拍值，不推 0 / Fault: output frozen, never zeroed *)
        tBadElapsed := tonBad.ET;
        bValid      := FALSE;

    ELSE
        eState    := eFault;
        bValid    := FALSE;
        bHolding  := FALSE;
        bTimedOut := FALSE;
        uErrorId  := 16#0007_0005;                 // 故障级：非法状态 / Fault: illegal state

END_CASE;

(* —— 段 7：出口映射（bError 与 uErrorId 同源；bTimedOut 为信息级不置 bError） —— *)
bError := (uErrorId <> 16#0007_0000) AND (uErrorId <> 16#0007_0001);

END_FUNCTION_BLOCK
